// TwinCAT 3 PLC project IAG50cm
// ProjectVersion: 0.10.0
// ProgramVersion: 3.1.4026.12
// libraries:
//   BROTLib, 0.20.0 (BROT)
//   VisuElemBase, * (System)
//   VisuInputs, * (System)
//   Tc2_Math, * (Beckhoff Automation GmbH)
//   Tc2_MC2, * (Beckhoff Automation GmbH)
//   Tc2_MC2_Drive, * (Beckhoff Automation GmbH)
//   Tc2_SerialCom, * (Beckhoff Automation GmbH)
//   Tc2_Standard, * (Beckhoff Automation GmbH)
//   Tc2_System, * (Beckhoff Automation GmbH)
//   Tc2_Utilities, * (Beckhoff Automation GmbH)
//   Tc3_IotBase, * (Beckhoff Automation GmbH)
//   Tc3_IotCommunicator, * (Beckhoff Automation GmbH)
//   Tc3_MC2_AdvancedHoming, * (Beckhoff Automation GmbH)
//   Tc3_Module, * (Beckhoff Automation GmbH)
//   VisuDialogs, * (System)
//   AstroBROT,0.4.3,BROT
//   VisuSymbols,newest,System
// project tree:
//   DUTs/ E_MirrorCoverState.TcDUT, ST_AxisStatus.TcDUT
//   / GlobalTextList.TcGTLO, PlcTask.TcTTO, PlcTask_Fast.TcTTO, Visualization Manager.TcVMO (not stored)
//   GVLs/ GVL_Homing.TcGVL, GVL_Pointing.TcGVL, GVL_Safety.TcGVL, GVL_Serial.TcGVL, Global_Version.TcGVL
//   POUs/CoverControl/ FB_CoverControl.TcPOU
//   POUs/CoverControl/States/ FB_CoverClosingState.TcPOU, FB_CoverIdleState.TcPOU, FB_CoverOpeningState.TcPOU, FB_CoverState.TcPOU, FB_CoverStoppingState.TcPOU, I_CoverState.TcIO
//   POUs/DomeControl/ FB_DomeControl.TcPOU
//   POUs/DomeControl/States/ FB_DomeClosingState.TcPOU, FB_DomeErrorState.TcPOU, FB_DomeHomingState.TcPOU, FB_DomeIdleState.TcPOU, FB_DomeOpeningState.TcPOU, FB_DomeParkingState.TcPOU, FB_DomeStoppingState.TcPOU, FB_DomeState.TcPOU, FB_DomeMovingState.TcPOU, I_DomeState.TcIO
//   POUs/ FB_LatchHome.TcPOU, FB_SafetyHandling.TcPOU, FB_SerialBackground.TcPOU, FB_HomeDropReason.TcPOU, FB_HomeHold.TcPOU, FB_StartRequest.TcPOU, FB_StepDrain.TcPOU, FB_SweepStop.TcPOU, SerialBackground.TcPOU, FB_AxisControl.TcPOU, FB_CabinetControl.TcPOU, FB_FocusControl.TcPOU, FB_HourAngleControl.TcPOU, FB_DeclinationControl.TcPOU, FB_TelescopeControl.TcPOU, MAIN.TcPOU
//   POUs/Functions/ F_HourAngleOffsetOnAxis.TcPOU, F_RoundLREAL.TcPOU, NCError_TO_STRING.TcPOU
//   POUs/PendantControl/ FB_PendantControl.TcPOU
//   POUs/PendantControl/States/ FB_PendantErrorState.TcPOU, FB_PendantPreInitState.TcPOU, FB_PendantSetDECState.TcPOU, FB_PendantSetFocusState.TcPOU, FB_PendantSetHAState.TcPOU, FB_PendantInitState.TcPOU, FB_PendantState.TcPOU, FB_PendantIdleState.TcPOU, I_PendantState.TcIO
//   POUs/Pointing/ FB_PointingModelForward.TcPOU, FB_PointingModelInversion.TcPOU
//   POUs/Testing/ FB_RefMarkerSearch.TcPOU
//   VISUs/ Safety.TcVIS
// real-time tasks:
//   TASK PlcTask: cycle T#10ms, priority 20, ADS port 350
//   TASK VISU_TASK: cycle T#200000us, priority 30, ADS port 351
//   TASK PlcTask_Fast: cycle T#2ms, priority 19, ADS port 352
// motion (NC):
//   TASK NC-Task 1 SAF: cycle T#2ms, priority 4, ADS port 501
//   TASK NC-Task 1 SVB: cycle T#10ms, priority 8, ADS port 511
//   AXIS Declination (id 1)
//     General: UnitName=°
//     Dynamic: Acceleration=3.21148, Deceleration=3.21148, Jerk=4.13844
//     Velo: RefSearch=0.10384, RefSync=0.10384, SlowManual=0.5192, FastManual=3.1152, Fast=10.384, Maximum=10.384
//     TargetPosControl: Range=0.5
//     OtherSettings: AllowMotionCmdToSlave=true
//     encoder EncType=4
//       EncPara: ScaleFactorNumerator=360, ScaleFactorDenominator=36864000, Offset=-23, Inverse=true, MaxCount=#xffffffff
//         Inc: RefMode=2
//     drive DrvType=16
//       DrvPara: MaxCount=#xffffffff, DriveControlDWord=#x00020000
//         Analog: VeloReferenz=11.4224, VeloScale=312, TorqueSetpointScale=10, ScaleFactorActTorque=0.1
//         TimeComp: TaskDelayCycles=1
//     controller CtrType=1
//       CtrPara: PriorControlFactor=1
//         PID: PosKp=3
//         Observer: BandWidth=20
//   AXIS HourAngle (id 2)
//     General: UnitName=°
//     Dynamic: Acceleration=3.6, Deceleration=3.6, Jerk=3.19705
//     Velo: RefSearch=0.10384, RefSync=0.10384, SlowManual=0.5192, FastManual=3.1152, Fast=10.384, Maximum=10.384
//     TargetPosControl: Range=0.5
//     OtherSettings: AllowMotionCmdToSlave=true
//     encoder EncType=4
//       EncPara: ScaleFactorNumerator=360, ScaleFactorDenominator=36864000, Inverse=true, MaxCount=#xffffffff
//         Inc: RefMode=2
//     drive DrvType=16
//       DrvPara: MaxCount=#xffffffff, DriveControlDWord=#x00020000
//         Analog: VeloReferenz=11.4224, VeloScale=312, TorqueSetpointScale=10, ScaleFactorActTorque=0.1
//         TimeComp: TaskDelayCycles=1
//     controller CtrType=1
//       CtrPara: PriorControlFactor=1
//         Observer: BandWidth=20
//   AXIS Focus (id 3)
//     Dynamic: AccelerationMaximum=15, DecelerationMaximum=15, Acceleration=1, Deceleration=1, Jerk=10
//     Velo: RefSearch=0.26997, RefSync=0.26997, SlowManual=0.1, FastManual=1, Fast=26.997, Maximum=2
//     OtherSettings: AllowMotionCmdToSlave=true, PulseDistancePos=1, PulseDistanceNeg=1
//     encoder EncType=19
//       EncPara: ScaleFactorNumerator=3, ScaleFactorDenominator=10485760, Offset=9.78274383544922, MaxCount=#xffffffff, ReferenceSystem=1
//         SoftEndMinControl: Enable=true, Range=1
//         SoftEndMaxControl: Enable=true, Range=17
//     drive DrvType=16
//       DrvPara: MaxCount=#xffffffff, DriveControlDWord=#x00020100
//         Analog: VeloReferenz=29.6967, VeloScale=32, TorqueSetpointScale=10, ScaleFactorActTorque=0.1
//         TimeComp: TaskDelayCycles=1
//     controller CtrType=1
//       CtrPara: PriorControlFactor=1
//         Observer: BandWidth=20
// I/O:
//   DEVICE Device 1 (EtherCAT), AmsNetId 5.146.183.126.2.1
//     Term 1 (EK1200) [EK1200-5000 EtherCAT Power supply (2A E-Bus)]
//       Safety (EL1918) [EL1918, 8Ch. Safety Input 24V, TwinSAFE]
//         modules: Module 2 (FSLOGIC)
//       Safety Out (EL2904) [EL2904, 4 Ch. Safety Output 24V, 0.5A, TwinSAFE]
//         modules: Module 1 (FSOES), Module 2 (DO)
//       Power Status (EL1808) [EL1808 8Ch. Dig. Input 24V, 3ms]
//       HA DEC (ELM7212-9016) [ELM7212-9016 2Ch. Servo Terminal (48 V, 4,5 A RMS, OCT, STO, TwinSAFE Logic)]
//         modules: Module 1 (SAFETY)
//         startup 32785:21 := 0E01 // DRV Motor Settings Ch.1 / Commutation offset
//         startup 32785:27 := 10270000 // DRV Motor Settings Ch.1 / Motor speed limitation
//         startup 32786:19 := 0000 // DRV Brake Settings Ch.1 / Emergency application timeout
//         startup 32784:51 := 0A00 // DRV Amplifier Settings Ch.1 / Stand still window
//         startup 28688:11 := F90C // DRV Outputs Ch.1 / Torque limitation
//         startup 32784:19 := FD00 // DRV Amplifier Settings Ch.1 / Current loop proportional gain
//         startup 32784:18 := 0600 // DRV Amplifier Settings Ch.1 / Current loop integral time
//         startup 32784:21 := 48000000 // DRV Amplifier Settings Ch.1 / Velocity loop proportional gain
//         startup 32784:20 := 96000000 // DRV Amplifier Settings Ch.1 / Velocity loop integral time
//         startup 33041:21 := 0E01 // DRV Motor Settings Ch.2 / Commutation offset
//         startup 33041:27 := 10270000 // DRV Motor Settings Ch.2 / Motor speed limitation
//         startup 33042:19 := 0000 // DRV Brake Settings Ch.2 / Emergency application timeout
//         startup 33040:51 := 0A00 // DRV Amplifier Settings Ch.2 / Stand still window
//         startup 28944:11 := F90C // DRV Outputs Ch.2 / Torque limitation
//         startup 33040:19 := FD00 // DRV Amplifier Settings Ch.2 / Current loop proportional gain
//         startup 33040:18 := 0600 // DRV Amplifier Settings Ch.2 / Current loop integral time
//         startup 33040:21 := 48000000 // DRV Amplifier Settings Ch.2 / Velocity loop proportional gain
//         startup 33040:20 := 96000000 // DRV Amplifier Settings Ch.2 / Velocity loop integral time
//       MirrorCover1 (EL2652) [EL2652 2Ch. Relay Output, CO (230V AC / 30V DC)]
//       MirrorCover2 (EL2652) [EL2652 2Ch. Relay Output, CO (230V AC / 30V DC)]
//       Power (EL9110) [EL9110 Power Supplier with LED (24V, Diagnostics)]
//       Reset 24V (EL2004) [EL2004 4Ch. Dig. Output 24V, 0.5A]
//       FOCUS (ELM7221-9016) [ELM7221-9016 1Ch. Servo Terminal (48 V, 8 A RMS, OCT, STO, TwinSAFE Logic)]
//         modules: Module 1 (SAFETY)
//         startup 32785:21 := 0E01 // DRV Motor Settings Ch.1 / Commutation offset
//         startup 32785:27 := 10270000 // DRV Motor Settings Ch.1 / Motor speed limitation
//         startup 32786:19 := 0000 // DRV Brake Settings Ch.1 / Emergency application timeout
//         startup 32784:51 := 0A00 // DRV Amplifier Settings Ch.1 / Stand still window
//         startup 28688:11 := FC0D // DRV Outputs Ch.1 / Torque limitation
//         startup 32784:19 := FD00 // DRV Amplifier Settings Ch.1 / Current loop proportional gain
//         startup 32784:18 := 0600 // DRV Amplifier Settings Ch.1 / Current loop integral time
//         startup 32784:21 := 47000000 // DRV Amplifier Settings Ch.1 / Velocity loop proportional gain
//         startup 32784:20 := 96000000 // DRV Amplifier Settings Ch.1 / Velocity loop integral time
//       Encoder DEC (EL5021) [EL5021 1Ch. Sin/Cos Encoder]
//       Encoder HA (EL5021) [EL5021 1Ch. Sin/Cos Encoder]
//       Cabinet IN (EL1004) [EL1004 4Ch. Dig. Input 24V, 3ms]
//       Dome Pendant (EL6002) [EL6002 Interface 2Ch. (RS232)]
//       Term 13 (EL9011) [EL9011 End Terminal]
// variable links:
//   Device 1 (EtherCAT) <-> Device 1 (EtherCAT)/Term 1 (EK1200)/FOCUS (ELM7221-9016)
//     Term 1 (EK1200)/Safety (EL1918)/ConnectionOutputs/TwinSafeGroup1.Connection to Term 12 (ELM7221-9016)_3 RxPDO <-> Module 1 (SAFETY)/SAFETY FSoE Connection 1 Send Message/Message_1
//   Device 1 (EtherCAT) <-> Device 1 (EtherCAT)/Term 1 (EK1200)/HA DEC (ELM7212-9016)
//     Term 1 (EK1200)/Safety (EL1918)/ConnectionInputs/TwinSafeGroup1.Connection to Term 4 (ELM7212-9016)_4 TxPDO <-> Module 1 (SAFETY)/SAFETY FSoE Connection 1 Receive Message/Message_1
//     Term 1 (EK1200)/Safety (EL1918)/ConnectionOutputs/TwinSafeGroup1.Connection to Term 4 (ELM7212-9016)_4 RxPDO <-> Module 1 (SAFETY)/SAFETY FSoE Connection 1 Send Message/Message_1
//   Device 1 (EtherCAT) <-> Device 1 (EtherCAT)/Term 1 (EK1200)/Safety (EL1918)
//     Term 1 (EK1200)/FOCUS (ELM7221-9016)/Module 1 (SAFETY)/SAFETY FSoE Connection 1 Receive Message/Message_1 <-> ConnectionInputs/TwinSafeGroup1.Connection to Term 12 (ELM7221-9016)_3 TxPDO
//     Term 1 (EK1200)/Safety Out (EL2904)/Module 1 (FSOES)/RxPDO/FSOE <-> ConnectionInputs/TwinSafeGroup1.EL2904, 4 digital outputs_1_7 TxPDO
//   Device 1 (EtherCAT) <-> Device 1 (EtherCAT)/Term 1 (EK1200)/Safety Out (EL2904)
//     Term 1 (EK1200)/Safety (EL1918)/ConnectionOutputs/TwinSafeGroup1.EL2904, 4 digital outputs_1_7 RxPDO <-> Module 1 (FSOES)/TxPDO/FSOE
//   NC-Task 1 SAF/Axes/Declination <-> Device 1 (EtherCAT)/Term 1 (EK1200)/Encoder DEC (EL5021)
//     Enc/Inputs/In/nDataIn1 <-> ENC Status/Counter value
//     Enc/Inputs/In/nDataIn2 <-> ENC Status/Latch value
//     Enc/Inputs/In/nDcInputTime <-> InfoData/DcInputShift
//     Enc/Inputs/In/nState1 <-> ENC Status/Latch C valid
//     Enc/Inputs/In/nState1 @bit 2 <-> ENC Status/Set counter done
//     Enc/Inputs/In/nState2 @bit 2 <-> ENC Status/Status of input C
//     Enc/Inputs/In/nState2 @bit 5 <-> ENC Status/Sync error
//     Enc/Inputs/In/nState2 @bit 6 <-> ENC Status/TxPDO State
//     Enc/Inputs/In/nState2 @bit 7 <-> ENC Status/TxPDO Toggle
//     Enc/Inputs/In/nState3 @bit 4 <-> ENC Status/Amplitude error
//     Enc/Inputs/In/nState3 @bit 3 <-> ENC Status/Frequency error
//     Enc/Inputs/In/nState4 @bit 1 <-> WcState/InputToggle
//     Enc/Inputs/In/nState4 <-> WcState/WcState
//     Enc/Outputs/Out/nCtrl1 @bit 1 <-> ENC Control/Enable latch C
//     Enc/Outputs/Out/nCtrl1 @bit 2 <-> ENC Control/Set counter
//     Enc/Outputs/Out/nDataOut1 <-> ENC Control/Set counter value
//   NC-Task 1 SAF/Axes/Declination <-> Device 1 (EtherCAT)/Term 1 (EK1200)/HA DEC (ELM7212-9016)
//     Drive/Inputs/In/nDcOutputTime <-> InfoData/DcOutputShift
//     Drive/Inputs/In/nState1 <-> DRV Statusword Channel 1/Statusword
//     Drive/Inputs/In/nState2 <-> DRV Statusword Channel 1/Statusword @bit 8
//     Drive/Inputs/In/nState4 @bit 1 <-> WcState/InputToggle0
//     Drive/Inputs/In/nState4 <-> WcState/WcState0
//     Drive/Outputs/Out/nCtrl1 <-> DRV Controlword Channel 1/Controlword
//     Drive/Outputs/Out/nCtrl2 <-> DRV Controlword Channel 1/Controlword @bit 8
//     Drive/Outputs/Out/nDataOut2 <-> DRV Target velocity Channel 1/Target velocity
//   NC-Task 1 SAF/Axes/Focus <-> Device 1 (EtherCAT)/Term 1 (EK1200)/FOCUS (ELM7221-9016)
//     Drive/Inputs/In/nDataIn1 <-> DRV Following error actual value/Following error actual value
//     Drive/Inputs/In/nDcOutputTime <-> InfoData/DcOutputShift
//     Drive/Inputs/In/nState1 <-> DRV Statusword/Statusword
//     Drive/Inputs/In/nState2 <-> DRV Statusword/Statusword @bit 8
//     Drive/Inputs/In/nState4 @bit 1 <-> WcState/InputToggle0
//     Drive/Inputs/In/nState4 <-> WcState/WcState0
//     Drive/Outputs/Out/nCtrl1 <-> DRV Controlword/Controlword
//     Drive/Outputs/Out/nCtrl2 <-> DRV Controlword/Controlword @bit 8
//     Drive/Outputs/Out/nDataOut1 <-> DRV Target position/Target position
//     Enc/Inputs/In/nDataIn1 <-> FB Position/Position
//     Enc/Inputs/In/nDcInputTime <-> InfoData/DcInputShift
//     Enc/Inputs/In/nState4 @bit 1 <-> WcState/InputToggle0
//     Enc/Inputs/In/nState4 <-> WcState/WcState0
//   NC-Task 1 SAF/Axes/HourAngle <-> Device 1 (EtherCAT)/Term 1 (EK1200)/Encoder HA (EL5021)
//     Enc/Inputs/In/nDataIn1 <-> ENC Status/Counter value
//     Enc/Inputs/In/nDataIn2 <-> ENC Status/Latch value
//     Enc/Inputs/In/nState1 <-> ENC Status/Latch C valid
//     Enc/Inputs/In/nState1 @bit 2 <-> ENC Status/Set counter done
//     Enc/Inputs/In/nState2 @bit 2 <-> ENC Status/Status of input C
//     Enc/Inputs/In/nState2 @bit 5 <-> ENC Status/Sync error
//     Enc/Inputs/In/nState2 @bit 6 <-> ENC Status/TxPDO State
//     Enc/Inputs/In/nState2 @bit 7 <-> ENC Status/TxPDO Toggle
//     Enc/Inputs/In/nState3 @bit 4 <-> ENC Status/Amplitude error
//     Enc/Inputs/In/nState3 @bit 3 <-> ENC Status/Frequency error
//     Enc/Inputs/In/nState4 @bit 1 <-> WcState/InputToggle
//     Enc/Inputs/In/nState4 <-> WcState/WcState
//     Enc/Outputs/Out/nCtrl1 @bit 1 <-> ENC Control/Enable latch C
//     Enc/Outputs/Out/nCtrl1 @bit 2 <-> ENC Control/Set counter
//     Enc/Outputs/Out/nDataOut1 <-> ENC Control/Set counter value
//   NC-Task 1 SAF/Axes/HourAngle <-> Device 1 (EtherCAT)/Term 1 (EK1200)/HA DEC (ELM7212-9016)
//     Drive/Inputs/In/nDcOutputTime <-> InfoData/DcOutputShift
//     Drive/Inputs/In/nState1 <-> DRV Statusword Channel 2/Statusword
//     Drive/Inputs/In/nState2 <-> DRV Statusword Channel 2/Statusword @bit 8
//     Drive/Inputs/In/nState4 @bit 1 <-> WcState/InputToggle0
//     Drive/Inputs/In/nState4 <-> WcState/WcState0
//     Drive/Outputs/Out/nCtrl1 <-> DRV Controlword Channel 2/Controlword
//     Drive/Outputs/Out/nCtrl2 <-> DRV Controlword Channel 2/Controlword @bit 8
//     Drive/Outputs/Out/nDataOut2 <-> DRV Target velocity Channel 2/Target velocity
//   IAG50cm/IAG50cm Instance <-> Device 1 (EtherCAT)/Term 1 (EK1200)/Cabinet IN (EL1004)
//     PlcTask Inputs/MAIN.telescopeControl.fbCabinet.bIMode <-> Channel 1/MAIN.telescopeControl.fbCabinet.bIMode
//     PlcTask Inputs/MAIN.telescopeControl.fbCabinet.bIReset <-> Channel 2/MAIN.telescopeControl.fbCabinet.bIReset
//   IAG50cm/IAG50cm Instance <-> Device 1 (EtherCAT)/Term 1 (EK1200)/Dome Pendant (EL6002)
//     PlcTask_Fast Inputs/SerialBackground.fbDomeSerial.stIn_EL6001/D <-> COM TxPDO-Map Inputs Channel 2/Data In 0
//     PlcTask_Fast Inputs/SerialBackground.fbDomeSerial.stIn_EL6001/D @bit {8..168 step 8} <-> COM TxPDO-Map Inputs Channel 2/Data In {1..21}  (21 links)
//     PlcTask_Fast Inputs/SerialBackground.fbDomeSerial.stIn_EL6001/Status <-> COM TxPDO-Map Inputs Channel 2/Status
//     PlcTask_Fast Inputs/SerialBackground.fbPendantSerial.stIn_EL6001/D <-> COM TxPDO-Map Inputs Channel 1/Data In 0
//     PlcTask_Fast Inputs/SerialBackground.fbPendantSerial.stIn_EL6001/D @bit {8..168 step 8} <-> COM TxPDO-Map Inputs Channel 1/Data In {1..21}  (21 links)
//     PlcTask_Fast Inputs/SerialBackground.fbPendantSerial.stIn_EL6001/Status <-> COM TxPDO-Map Inputs Channel 1/Status
//     PlcTask_Fast Outputs/SerialBackground.fbDomeSerial.stOut_EL6001/Ctrl <-> COM RxPDO-Map Outputs Channel 2/Ctrl
//     PlcTask_Fast Outputs/SerialBackground.fbDomeSerial.stOut_EL6001/D <-> COM RxPDO-Map Outputs Channel 2/Data Out 0
//     PlcTask_Fast Outputs/SerialBackground.fbDomeSerial.stOut_EL6001/D @bit {8..168 step 8} <-> COM RxPDO-Map Outputs Channel 2/Data Out {1..21}  (21 links)
//     PlcTask_Fast Outputs/SerialBackground.fbPendantSerial.stOut_EL6001/Ctrl <-> COM RxPDO-Map Outputs Channel 1/Ctrl
//     PlcTask_Fast Outputs/SerialBackground.fbPendantSerial.stOut_EL6001/D <-> COM RxPDO-Map Outputs Channel 1/Data Out 0
//     PlcTask_Fast Outputs/SerialBackground.fbPendantSerial.stOut_EL6001/D @bit {8..168 step 8} <-> COM RxPDO-Map Outputs Channel 1/Data Out {1..21}  (21 links)
//   IAG50cm/IAG50cm Instance <-> Device 1 (EtherCAT)/Term 1 (EK1200)/FOCUS (ELM7221-9016)
//     PlcTask Outputs/GVL_Safety.ErrAck <-> Module 1 (SAFETY)/SAFETY Standard Outputdata/Standard In Var 3
//     PlcTask Outputs/GVL_Safety.Run <-> Module 1 (SAFETY)/SAFETY Standard Outputdata/Standard In Var 2
//   IAG50cm/IAG50cm Instance <-> Device 1 (EtherCAT)/Term 1 (EK1200)/HA DEC (ELM7212-9016)
//     PlcTask Outputs/GVL_Safety.ErrAck <-> Module 1 (SAFETY)/SAFETY Standard Outputdata/Standard In Var 3
//     PlcTask Outputs/GVL_Safety.Run <-> Module 1 (SAFETY)/SAFETY Standard Outputdata/Standard In Var 2
//   IAG50cm/IAG50cm Instance <-> Device 1 (EtherCAT)/Term 1 (EK1200)/MirrorCover1 (EL2652)
//     PlcTask Outputs/MAIN.coverControl.bMotor1RelaisA <-> Channel 1/Output
//     PlcTask Outputs/MAIN.coverControl.bMotor1RelaisB <-> Channel 2/Output
//   IAG50cm/IAG50cm Instance <-> Device 1 (EtherCAT)/Term 1 (EK1200)/MirrorCover2 (EL2652)
//     PlcTask Outputs/MAIN.coverControl.bMotor2RelaisA <-> Channel 1/Output
//     PlcTask Outputs/MAIN.coverControl.bMotor2RelaisB <-> Channel 2/Output
//   IAG50cm/IAG50cm Instance <-> Device 1 (EtherCAT)/Term 1 (EK1200)/Power Status (EL1808)
//     PlcTask Inputs/MAIN.telescopeControl.fbCabinet.bAuxiliaryContact24V <-> Channel 1/Input
//     PlcTask Inputs/MAIN.telescopeControl.fbCabinet.bAuxiliaryContact48V <-> Channel 2/Input
//     PlcTask Inputs/MAIN.telescopeControl.fbCabinet.bAuxiliaryContactFOCUS <-> Channel 4/Input
//     PlcTask Inputs/MAIN.telescopeControl.fbCabinet.bAuxiliaryContactHADEC <-> Channel 3/Input
//     PlcTask Inputs/MAIN.telescopeControl.fbCabinet.bCollectiveReport24VFuse <-> Channel 6/Input
//     PlcTask Inputs/MAIN.telescopeControl.fbCabinet.bState24VFuse <-> Channel 5/Input
//   IAG50cm/IAG50cm Instance <-> Device 1 (EtherCAT)/Term 1 (EK1200)/Reset 24V (EL2004)
//     PlcTask Outputs/MAIN.telescopeControl.fbCabinet.bOErrorLED <-> Channel 2/MAIN.telescopeControl.fbCabinet.bOErrorLED
//   IAG50cm/IAG50cm Instance <-> Device 1 (EtherCAT)/Term 1 (EK1200)/Safety (EL1918)
//     PlcTask Inputs/MAIN.safetyHandling.stInfoEStop1 <-> Function Block Info Data/TwinSafeGroup1.SS1.FBMon1 Info Data
//     PlcTask Inputs/MAIN.safetyHandling.stInfoGroup1 <-> TwinSAFE Group Info Data/TwinSafeGroup1 Info Data
//     PlcTask Outputs/GVL_Safety.ErrAck <-> StandardOutputs/TwinSafeGroup1.ErrorAcknowledgement_2
//     PlcTask Outputs/GVL_Safety.Restart <-> StandardOutputs/TwinSafeGroup1.Restart_6
//     PlcTask Outputs/GVL_Safety.Run <-> StandardOutputs/TwinSafeGroup1.Run_1
//   IAG50cm/IAG50cm Instance <-> NC-Task 1 SAF/Axes/Declination
//     PlcTask Inputs/MAIN.decControl.axisRef.NcToPlc <-> Outputs/ToPlc
//     PlcTask Outputs/MAIN.decControl.axisRef.PlcToNc <-> Inputs/FromPlc
//   IAG50cm/IAG50cm Instance <-> NC-Task 1 SAF/Axes/Focus
//     PlcTask Inputs/MAIN.focusControl.axisRef.NcToPlc <-> Outputs/ToPlc
//     PlcTask Outputs/MAIN.focusControl.axisRef.PlcToNc <-> Inputs/FromPlc
//   IAG50cm/IAG50cm Instance <-> NC-Task 1 SAF/Axes/HourAngle
//     PlcTask Inputs/MAIN.haControl.axisRef.NcToPlc <-> Outputs/ToPlc
//     PlcTask Outputs/MAIN.haControl.axisRef.PlcToNc <-> Inputs/FromPlc

CONFIGURATION IAG50cm
    RESOURCE PLC ON TwinCAT3
        TASK PlcTask(INTERVAL := T#10ms, PRIORITY := 20);
        TASK PlcTask_Fast(INTERVAL := T#2ms, PRIORITY := 19);
        PROGRAM MAIN WITH PlcTask : MAIN;
        PROGRAM SerialBackground WITH PlcTask_Fast : SerialBackground;
    END_RESOURCE
END_CONFIGURATION

// ---- DUTs/E_MirrorCoverState.TcDUT
{attribute 'qualified_only'}
{attribute 'strict'}
//{attribute 'to_string'}
TYPE E_MirrorCoverState :
(
	closing := 0,
	opening := 1,
	stopped := 2,
	closed	:= 3,
	open	:= 4,
	error := 5,
	unknown := 6
);
END_TYPE

// ---- DUTs/ST_AxisStatus.TcDUT
// Plan step 3.2: the feedback of one axis (FB_Axis outputs) as read once per scan by FB_TelescopeControl._ReadAxes. Same struct as
// MONETcommon's (it moves to BROTLib in step 4). The axes' outputs do not change while the telescope body runs, so reading them into
// one struct is the same as reading fbAxis.* at every use.
TYPE ST_AxisStatus :
STRUCT
	bStandStill		: BOOL;
	bStopDone		: BOOL;
	bInMotion		: BOOL;
	bInRamp			: BOOL;
	bHoming			: BOOL;
	bStopping		: BOOL;
	bBusy			: BOOL;
	bTracking		: BOOL;
END_STRUCT
END_TYPE

// ---- GVLs/GVL_Homing.TcGVL
{attribute 'qualified_only'}
VAR_GLOBAL
	// #113: how FB_LatchHome ends the calibration sweep after a stop. Test switch, written over ADS (GVL_Homing.nAbortMode),
	// so the approaches can be tried one after the other without a new activation. Not persistent.
	//   0: as before (MC_AbortHoming into the running step: never completes, 4F000001 after 10 s)
	//   1: no MC_AbortHoming while a step block is Busy, the axis is reset instead (reset=1 clears HomingBusy)
	//   2: the Busy reference step keeps its Execute while MC_AbortHoming runs
	//   3: MC_AbortHoming with DisableDriveAccess FALSE
	nAbortMode		: INT := 1;
END_VAR

// ---- GVLs/GVL_Pointing.TcGVL
VAR_GLOBAL
	(* values of the pointing model
	Hour Angle	: tau
	Declination	: dec
	*)

	(*
	 pointing from: 21.01.2026 136 points (from Lukas Melzig)
	RMS Ha:  17.69244750276253
	RMS Dec:  13.468555776826959
	*)
	C_mAl_tau	: LREAL := 0.01687078;
	C_mEl_tau	: LREAL := -0.02608578;
	C_Coll_tau	: LREAL := 0.29826615;
	C_Refr_tau	: LREAL := -0.00759962;
	C_Enc_tau	: LREAL := 0.00108764;
	C_Flex_tau	: LREAL := -0.02462705;
	C_NP_tau	: LREAL := 0.02128217;
	
	C_mAl_dec	: LREAL := 0.01606325;
	C_mEl_dec	: LREAL := -0.05749048;
	C_Coll_dec	: LREAL := -0.17376101;
	C_Refr_dec	: LREAL := 0.01678090;
	C_Flex_dec	: LREAL := -0.01915146;
END_VAR

// ---- GVLs/GVL_Safety.TcGVL
{attribute 'qualified_only'}
VAR_GLOBAL
	// Run/Stop Safety
	Run			AT%Q*:	BOOL;
	// Restart Safety
	Restart		AT%Q*:	BOOL;
	// Error Acknowledgement 
	ErrAck		AT%Q*:	BOOL;

END_VAR

// ---- GVLs/GVL_Serial.TcGVL
VAR_GLOBAL
	RxBufferDome			: ComBuffer;	(* Receive data buffer; used with all receive function blocks *)
	TxBufferDome			: ComBuffer;	(* Transmit data buffer; used with all receive function blocks *)
	
	RxBufferPendant			: ComBuffer;	(* Receive data buffer; used with all receive function blocks *)
	TxBufferPendant			: ComBuffer;	(* Transmit data buffer; used with all receive function blocks *)
END_VAR

// ---- GVLs/Global_Version.TcGVL
{attribute 'qualified_only'}
VAR_GLOBAL CONSTANT
	// Mirrors Beckhoff's own Global_Version.stLibVersion_* pattern (see ST_LibVersion),
	// which only covers Tc2_*/Tc3_* library references, not custom ones -- until now: this
	// GVL uses Beckhoff's own naming exactly, so it merges into a consumer's Global_Version.
	// Kept in sync with <ProjectVersion> in IAG50cm.plcproj at release time.
	stLibVersion_IAG50cm : ST_LibVersion := (
		iMajor := 0,
		iMinor := 10,
		iBuild := 0,
		iRevision := 0,
		nFlags := 1,
		sVersion := '0.10.0'
	);
END_VAR

// ---- POUs/CoverControl/States/I_CoverState.TcIO
INTERFACE I_CoverState

METHOD CloseCommand : BOOL
VAR_INPUT
END_VAR
END_METHOD

METHOD OpenCommand : BOOL
VAR_INPUT
END_VAR
END_METHOD

METHOD RunState : BOOL
VAR_INPUT
END_VAR
END_METHOD

METHOD StopCommand : BOOL
VAR_INPUT
END_VAR
END_METHOD

METHOD SuccessfulFinished : BOOL
VAR_INPUT
END_VAR
END_METHOD

END_INTERFACE

// ---- POUs/DomeControl/States/I_DomeState.TcIO
INTERFACE I_DomeState


METHOD CloseCommand : BOOL
END_METHOD


METHOD FoundError : BOOL
END_METHOD


METHOD HomeCommand : BOOL
END_METHOD


METHOD MoveCommand : BOOL
END_METHOD


METHOD OpenCommand : BOOL
END_METHOD


METHOD ParkCommand : BOOL
END_METHOD


METHOD ResetCommand : BOOL
END_METHOD

METHOD RunState : BOOL
VAR_INPUT
END_VAR
END_METHOD


PROPERTY StateID : STRING
GET
END_GET
END_PROPERTY


METHOD StopCommand : BOOL
END_METHOD


METHOD SuccessfulFinished : BOOL
END_METHOD

END_INTERFACE

// ---- POUs/PendantControl/States/I_PendantState.TcIO
INTERFACE I_PendantState

METHOD DecCommand : BOOL
VAR_INPUT
END_VAR
END_METHOD

METHOD FocusCommand : BOOL
VAR_INPUT
END_VAR
END_METHOD

METHOD FoundError : BOOL
VAR_INPUT
END_VAR
END_METHOD

METHOD HaCommand : BOOL
VAR_INPUT
END_VAR
END_METHOD

METHOD InitCommand : BOOL
VAR_INPUT
END_VAR
END_METHOD

METHOD ResetCommand : BOOL
VAR_INPUT
END_VAR
END_METHOD

METHOD RunState : BOOL
VAR_INPUT
END_VAR
END_METHOD

PROPERTY StateID : STRING
GET
END_GET
END_PROPERTY

METHOD Timeout : BOOL
VAR_INPUT
END_VAR
END_METHOD

METHOD ToIdle : BOOL
VAR_INPUT
END_VAR
END_METHOD

END_INTERFACE

// ---- POUs/MAIN.TcPOU
PROGRAM MAIN
VAR
	comm			: FB_Comm_MQTT_Influx;
	coverControl	: FB_CoverControl(comm := comm);
	focusControl	: FB_FocusControl(comm:=comm);
	haControl		: FB_HourAngleControl(comm:=comm);
	decControl		: FB_DeclinationControl(comm:=comm);
	telescopeControl: FB_TelescopeControl(comm := comm);
	domeControl		: FB_DomeControl(comm := comm);
	pendantControl 	: FB_PendantControl(comm:=comm);
	safetyHandling	: FB_SafetyHandling(comm:=comm);
	rtrigStartUpDone: R_TRIG;
	//search			: FB_RefMarkerSearch(); // use for searching for the Heideinhain encoder reference markers

	
END_VAR
VAR CONSTANT
	telescopeConfig		: ST_TelescopeConfig := (longitude := 9.9452433, latitude := 51.5592378, altitude := 100.0, 
													houranglePark := 0.0, declinationPark := 52.0, focusPark:= 16.3,
													hourangleHome := 0.0, declinationHome := 52.0, focusHome:= 16.3,
													name := 'Emmy Noether', diameter := 0.5, cabinet := 'Beckhoff', manufacturer := '???',
													mountOptions := 'HA-DEC', mount := 'HA_DEC');
END_VAR

//search(Enable:=TRUE); // use for reference marker search

domeControl(ipTelescope	:= telescopeControl);

pendantControl(
	ipTelescope	:= telescopeControl,
	ipFocus		:= focusControl);

coverControl(
	Delta := T#5S,
	TimeToCycle := T#15S,
	bEmergency := safetyHandling.estop);	// previous cycle's value, see bEstopTriggered below (#15)
	
focusControl(
	fVelocity:=1);
	
haControl();
decControl();
telescopeControl(
	fbHourAngle		:= haControl,
	fbDeclination	:= decControl,
	fbFocus			:= focusControl,
	fbDome			:= domeControl,
	fbCovers		:= coverControl,
	telescopeConfig	:= telescopeConfig,
	// was never wired, so STATUS.GLOBAL never reported the E-stop (BROTLib#10). safetyHandling runs below, so
	// this is the previous cycle's value; the drives are cut by the safety circuit regardless.
	bEstopTriggered	:= safetyHandling.estop,
	bSafetyAckPending	:= safetyHandling.ackPending,	// previous cycle, like bEstopTriggered (#59)
);

//Safety
// #11: a telescope reset (cabinet key or the reset command, only fires with an error or a pending acknowledge after an E-stop, #59) also gives the safety
// acknowledge, so the drives leave STO without the VISU
IF telescopeControl.bSafetyAckRequest THEN
	telescopeControl.bSafetyAckRequest := FALSE;
	safetyHandling.Acknowledge();
END_IF
safetyHandling();
// #103: one axis reset pass once the safety start-up is done (the start-up only acknowledges the drives)
rtrigStartUpDone(CLK := safetyHandling.bStartUpDone);
IF rtrigStartUpDone.Q THEN
	telescopeControl.bStartupAxisReset := TRUE;
END_IF

// Comm
comm(	
	sHostName			:= '169.254.149.100',
    nHostPort  			:= 1883,
    nKeepAlive  		:= 10,
	sTopicSub  		 	:= '50cm/Telescope/SET',
	sTopicPublish		:= '50cm/Telemetry',
	sTopicLog			:= '50cm/Log',
	Telescope			:= telescopeControl,
	RaDecTelescope		:= telescopeControl,
	Focus				:= focusControl,
	Dome				:= domeControl,
	MirrorCovers		:= coverControl,
);

END_PROGRAM

// ---- POUs/CoverControl/FB_CoverControl.TcPOU
FUNCTION_BLOCK FB_CoverControl IMPLEMENTS I_MirrorCovers
VAR_INPUT
	Delta		: TIME := T#5S;		// Time difference between both covers opening (and closing)
	TimeToCycle	: TIME := T#15S;	// Time for one motor to fully open/close
	// TRUE while the E-stop is triggered (MAIN: safetyHandling.estop): moving covers stop, open/close requests
	// are dropped (#15)
	bEmergency	: BOOL;
END_VAR
VAR_OUTPUT
END_VAR
VAR
	bOpen		: BOOL;
	bClose		: BOOL;
	bStop		: BOOL;
	// State
	fbCoverIdleState : FB_CoverIdleState(THIS);
	fbCoverOpeningState : FB_CoverOpeningState(THIS);
	fbCoverStoppingState : FB_CoverStoppingState(THIS);
	fbCoverClosingState : FB_CoverClosingState(THIS);
	
	ipState		: I_CoverState := fbCoverIdleState;
	// #111: the PLC cannot know the position of the covers after a start (activation, Reset Cold), so it starts with
	// "unknown" instead of assuming "closed". The first open or close cycle that completes sets the real end position.
	eCoverState	: E_MirrorCoverState := E_MirrorCoverState.unknown;
	// #71: TRUE only once an open or close cycle has completed since the PLC start. Until then the position is
	// unknown (the covers may be open after a restart), so a request is only ignored once the position is confirmed.
	bEndPositionConfirmed : BOOL := FALSE;
	bRequestIgnored : BOOL;
	// Trigger
	rtrigOpen		: R_TRIG;
	rtrigClose		: R_TRIG;
	rtrigStop		: R_TRIG;
	// Comm
	fbComm			: I_Comm;
	tonComm 		: TON := (PT:=T#5S);
	fbCoverOpenEvent:	FB_EventLog;
	fbCoverClosedEvent: FB_EventLog;
	fbCoverEmergencyEvent: FB_EventLog;
	fbCoverIgnoredEvent: FB_EventLog;
	// Motor relais
	bMotor1RelaisA	AT%Q*	: BOOL := FALSE;
	bMotor1RelaisB	AT%Q*	: BOOL := FALSE;
	
	bMotor2RelaisA	AT%Q*	: BOOL := FALSE;
	bMotor2RelaisB	AT%Q*	: BOOL := FALSE;
END_VAR

rtrigOpen(CLK := bOpen);
rtrigClose(CLK := bClose);
rtrigStop(CLK := bStop);
bRequestIgnored := FALSE;

IF bEmergency THEN
	// requests made during the E-stop are dropped (flags cleared below, #15)
	// stop only moving covers, so that closed/open covers keep their known state
	IF eCoverState = E_MirrorCoverState.opening OR eCoverState = E_MirrorCoverState.closing THEN
		ipState.StopCommand();
	END_IF
ELSE
	IF rtrigStop.Q THEN
		ipState.StopCommand();
	END_IF

	// #71: a request for the position the covers are confirmed to be in does nothing (it ran a full 20 s cycle)
	IF rtrigClose.Q THEN
		IF eCoverState = E_MirrorCoverState.closed AND bEndPositionConfirmed THEN
			bRequestIgnored := TRUE;
		ELSE
			ipState.CloseCommand();
		END_IF
	END_IF

	IF rtrigOpen.Q THEN
		IF eCoverState = E_MirrorCoverState.open AND bEndPositionConfirmed THEN
			bRequestIgnored := TRUE;
		ELSE
			ipState.OpenCommand();
		END_IF
	END_IF
END_IF

// #66: requests are one-shot. They are consumed in this scan whether they produced an edge or not, so a caller that
// repeats a request every scan (the park, stage 80) cannot leave a flag TRUE: left set, it would block the rising
// edge of every later request.
bOpen := FALSE;
bClose := FALSE;
bStop := FALSE;

ipState.RunState();

// send telemetry
tonComm(IN:=TRUE);
IF tonComm.Q THEN // publish new payload every second
	tonComm(IN:=FALSE);
	THIS^._SendTelemetry();	
END_IF


fbCoverOpenEvent(
	Trigger := eCoverState = E_MirrorCoverState.open,
	Level := ADSLOG_MSGTYPE_HINT,
	OnMessage := 'Mirror cover is open.',
	comm:= fbComm);
fbCoverClosedEvent(
	Trigger := eCoverState = E_MirrorCoverState.closed,
	Level := ADSLOG_MSGTYPE_HINT,
	OnMessage := 'Mirror cover is closed.',
	comm:= fbComm);
fbCoverIgnoredEvent(
	Trigger := bRequestIgnored,
	Level := ADSLOG_MSGTYPE_HINT,
	OnMessage := 'Mirror cover already in the requested end position, request ignored.',
	comm:= fbComm);
fbCoverEmergencyEvent(
	Trigger := bEmergency,
	Level := ADSLOG_MSGTYPE_WARN,
	OnMessage := 'Mirror cover: E-stop, covers stopped and commands ignored.',
	comm:= fbComm);

PROPERTY _CoverState : E_MirrorCoverState
SET
eCoverState := _CoverState;
bEndPositionConfirmed := (_CoverState = E_MirrorCoverState.closed OR _CoverState = E_MirrorCoverState.open);
END_SET
END_PROPERTY

PROPERTY _Motor1RelaisA : BOOL
SET
bMotor1RelaisA := _Motor1RelaisA;
END_SET
END_PROPERTY

PROPERTY _Motor1RelaisB : BOOL
SET
bMotor1RelaisB := _Motor1RelaisB;
END_SET
END_PROPERTY

PROPERTY _Motor2RelaisA : BOOL
SET
bMotor2RelaisA := _Motor2RelaisA;
END_SET
END_PROPERTY

PROPERTY _Motor2RelaisB : BOOL
SET
bMotor2RelaisB := _Motor2RelaisB;
END_SET
END_PROPERTY

METHOD _SendTelemetry : BOOL
VAR_INPUT
END_VAR
IF eCoverState = E_MirrorCoverState.closed THEN
	fbComm.PublishLREAL('telescope', 'dome', 'AUXILIARY.COVER.REALPOS', 0.0);
ELSIF eCoverState = E_MirrorCoverState.open THEN
	fbComm.PublishLREAL('telescope', 'dome', 'AUXILIARY.COVER.REALPOS', 1.0);
ELSE
	// moving, stopped or unknown (#111): not at an end position
	fbComm.PublishLREAL('telescope', 'dome', 'AUXILIARY.COVER.REALPOS', 0.5);
END_IF
END_METHOD

METHOD Close : BOOL
VAR_INPUT
END_VAR
bClose := TRUE;
END_METHOD

PROPERTY Closed : BOOL
GET
IF THIS^.CoverState = E_MirrorCoverState.closed THEN
	Closed := TRUE;
ELSE
	Closed := FALSE;
END_IF
END_GET
END_PROPERTY

PROPERTY CoverState : E_MirrorCoverState
GET
CoverState := eCoverState;
END_GET
END_PROPERTY

PROPERTY Error : BOOL
GET
Error := FALSE;
END_GET
END_PROPERTY

//FB_Init is always available implicitly and it is used primarily for initialization.
//The return value is not evaluated. For a specific influence, you can also declare the
//methods explicitly and provide additional code there with the standard initialization
//code. You can evaluate the return value.
METHOD FB_Init: BOOL
VAR_INPUT
    bInitRetains	: BOOL; // TRUE: the retain variables are initialized (reset warm / reset cold)
    bInCopyCode		: BOOL;  // TRUE: the instance will be copied to the copy code afterward (online change)
	comm			: I_Comm;
END_VAR
THIS^.fbComm 				:= comm;
END_METHOD

METHOD Open : BOOL
VAR_INPUT
END_VAR
bOpen := TRUE;
END_METHOD

PROPERTY Opened : BOOL
GET
IF THIS^.CoverState = E_MirrorCoverState.open THEN
	Opened := TRUE;
ELSE
	Opened := FALSE;
END_IF
END_GET
END_PROPERTY

METHOD Reset : BOOL
VAR_INPUT
END_VAR
END_METHOD

METHOD SetState : BOOL
VAR_INPUT
	newState :I_CoverState;
END_VAR
THIS^.ipState := newState;
END_METHOD

METHOD Stop : BOOL
VAR_INPUT
END_VAR
bStop := TRUE;
END_METHOD

END_FUNCTION_BLOCK

// ---- POUs/CoverControl/States/FB_CoverIdleState.TcPOU
FUNCTION_BLOCK FB_CoverIdleState EXTENDS FB_CoverState
VAR_INPUT
END_VAR
VAR_OUTPUT
END_VAR
VAR
END_VAR

METHOD CloseCommand : BOOL
pCover^.SetState(pCover^.fbCoverClosingState);
END_METHOD

METHOD OpenCommand : BOOL
pCover^.SetState(pCover^.fbCoverOpeningState);
END_METHOD

METHOD StopCommand : BOOL
pCover^.SetState(pCover^.fbCoverStoppingState);
END_METHOD

END_FUNCTION_BLOCK

// ---- POUs/CoverControl/States/FB_CoverState.TcPOU
FUNCTION_BLOCK FB_CoverState IMPLEMENTS I_CoverState
VAR_INPUT
END_VAR
VAR_OUTPUT
END_VAR
VAR
	pCover : POINTER TO FB_CoverControl;
END_VAR

{warning 'add method implementation '}
METHOD CloseCommand : BOOL
END_METHOD

METHOD FB_init : BOOL
VAR_INPUT
	bInitRetains : BOOL; // if TRUE, the retain variables are initialized (warm start / cold start)
	bInCopyCode : BOOL;  // if TRUE, the instance afterwards gets moved into the copy code (online change)
	pCover : POINTER TO FB_CoverControl;
END_VAR
THIS^.pCover := pCover;
END_METHOD

{warning 'add method implementation '}
METHOD OpenCommand : BOOL
END_METHOD

{warning 'add method implementation '}
METHOD RunState : BOOL
END_METHOD

{warning 'add method implementation '}
METHOD StopCommand : BOOL
END_METHOD

{warning 'add method implementation '}
METHOD SuccessfulFinished : BOOL
END_METHOD

END_FUNCTION_BLOCK

// ---- POUs/CoverControl/States/FB_CoverOpeningState.TcPOU
FUNCTION_BLOCK FB_CoverOpeningState EXTENDS FB_CoverState
VAR
	nStage			: UINT:= 0;
	tonDelta		: TON;		// PT is taken from pCover^.Delta at the start of each cycle (#76)
	tonFullCycle	: TON;		// PT is taken from pCover^.TimeToCycle at the start of each cycle (#76)
END_VAR

METHOD CloseCommand : BOOL
nStage := 0;
tonDelta(IN:=FALSE);
tonFullCycle(IN:=FALSE);
pCover^.SetState(pCover^.fbCoverClosingState);
END_METHOD

METHOD RunState : BOOL
tonDelta();
tonFullCycle();
CASE nStage OF
	0:
		// #76: the cycle times were only read once, by the declaration initialisers, so the inputs of FB_CoverControl
		// never reached the timers. Take them at the start of each cycle (not every scan: a change mid-cycle must not
		// end it early).
		tonDelta.PT := pCover^.Delta;
		IF pCover^.TimeToCycle > T#0S THEN
			tonFullCycle.PT := pCover^.TimeToCycle;
		ELSE
			tonFullCycle.PT := T#15S;	// 0 would declare the end position after one scan
		END_IF
		pCover^._CoverState := E_MirrorCoverState.opening;
		tonDelta.IN:=TRUE;
		nStage := 1;
	1:
		// Open Motor 1
		pCover^._Motor1RelaisA := TRUE;
		pCover^._Motor1RelaisB := FALSE;
		// Stop Motor 2
		pCover^._Motor2RelaisA := FALSE;
		pCover^._Motor2RelaisB := FALSE;
		nStage := 2;
	2:
		IF tonDelta.Q THEN
			tonDelta.IN:=FALSE;
			nStage:=3;
		END_IF 
	3:
		// Open Motor 2
		pCover^._Motor2RelaisA := TRUE;
		pCover^._Motor2RelaisB := FALSE;
		tonFullCycle.IN:=TRUE;
		nStage := 4;
	4:
		IF tonFullCycle.Q THEN
			tonFullCycle.IN:=FALSE;
			THIS^.SuccessfulFinished();
		END_IF 
END_CASE
END_METHOD

METHOD StopCommand : BOOL
nStage := 0;
tonDelta(IN:=FALSE);
tonFullCycle(IN:=FALSE);
pCover^.SetState(pCover^.fbCoverStoppingState);
END_METHOD

METHOD SuccessfulFinished : BOOL
nStage := 0;
tonDelta(IN:=FALSE);
tonFullCycle(IN:=FALSE);
// #71: release the relays at the end position (limit switches cut the motors, the covers are self-locking)
pCover^._Motor1RelaisA := FALSE;
pCover^._Motor1RelaisB := FALSE;
pCover^._Motor2RelaisA := FALSE;
pCover^._Motor2RelaisB := FALSE;
pCover^._CoverState := E_MirrorCoverState.open;
pCover^.SetState(pCover^.fbCoverIdleState);
END_METHOD

END_FUNCTION_BLOCK

// ---- POUs/CoverControl/States/FB_CoverStoppingState.TcPOU
FUNCTION_BLOCK FB_CoverStoppingState EXTENDS FB_CoverState
VAR_INPUT
END_VAR
VAR_OUTPUT
END_VAR
VAR
END_VAR

METHOD RunState : BOOL
// Stop Motor 1
pCover^._Motor1RelaisA := FALSE;
pCover^._Motor1RelaisB := FALSE;
// Stop Motor 2
pCover^._Motor2RelaisA := FALSE;
pCover^._Motor2RelaisB := FALSE;
THIS^.SuccessfulFinished();
END_METHOD

METHOD SuccessfulFinished : BOOL
pCover^._CoverState := E_MirrorCoverState.stopped;
pCover^.SetState(pCover^.fbCoverIdleState);
END_METHOD

END_FUNCTION_BLOCK

// ---- POUs/CoverControl/States/FB_CoverClosingState.TcPOU
FUNCTION_BLOCK FB_CoverClosingState EXTENDS FB_CoverState
VAR
	nStage			: UINT:= 0;
	tonDelta		: TON;		// PT is taken from pCover^.Delta at the start of each cycle (#76)
	tonFullCycle	: TON;		// PT is taken from pCover^.TimeToCycle at the start of each cycle (#76)
END_VAR

METHOD OpenCommand : BOOL
nStage := 0;
tonDelta(IN:=FALSE);
tonFullCycle(IN:=FALSE);
pCover^.SetState(pCover^.fbCoverOpeningState);
END_METHOD

METHOD RunState : BOOL
tonDelta();
tonFullCycle();
CASE nStage OF
	0:
		// #76: the cycle times were only read once, by the declaration initialisers, so the inputs of FB_CoverControl
		// never reached the timers. Take them at the start of each cycle (not every scan: a change mid-cycle must not
		// end it early).
		tonDelta.PT := pCover^.Delta;
		IF pCover^.TimeToCycle > T#0S THEN
			tonFullCycle.PT := pCover^.TimeToCycle;
		ELSE
			tonFullCycle.PT := T#15S;	// 0 would declare the end position after one scan
		END_IF
		pCover^._CoverState := E_MirrorCoverState.closing;
		tonDelta.IN := TRUE;
		nStage := 1;
	1:
		// Stop Motor 1
		pCover^._Motor1RelaisA := FALSE;
		pCover^._Motor1RelaisB := FALSE;
		// Close Motor 2
		pCover^._Motor2RelaisA := FALSE;
		pCover^._Motor2RelaisB := TRUE;
		nStage := 2;
	2:
		IF tonDelta.Q THEN
			tonDelta.IN := FALSE;
			nStage:=3;
		END_IF 
	3:
		// Close Motor 1
		pCover^._Motor1RelaisA := FALSE;
		pCover^._Motor1RelaisB := TRUE;
		tonFullCycle.IN:=TRUE;
		nStage := 4;
	4:
		IF tonFullCycle.Q THEN
			tonFullCycle.IN := FALSE;
			THIS^.SuccessfulFinished();
		END_IF 
END_CASE
END_METHOD

METHOD StopCommand : BOOL
nStage := 0;
tonDelta(IN:=FALSE);
tonFullCycle(IN:=FALSE);
pCover^.SetState(pCover^.fbCoverStoppingState);
END_METHOD

METHOD SuccessfulFinished : BOOL
nStage := 0;
tonDelta(IN:=FALSE);
tonFullCycle(IN:=FALSE);
// #71: release the relays at the end position (limit switches cut the motors, the covers are self-locking)
pCover^._Motor1RelaisA := FALSE;
pCover^._Motor1RelaisB := FALSE;
pCover^._Motor2RelaisA := FALSE;
pCover^._Motor2RelaisB := FALSE;
pCover^._CoverState := E_MirrorCoverState.closed;
pCover^.SetState(pCover^.fbCoverIdleState);
END_METHOD

END_FUNCTION_BLOCK

// ---- POUs/FB_FocusControl.TcPOU
FUNCTION_BLOCK FB_FocusControl EXTENDS FB_AxisControl IMPLEMENTS I_Focus
VAR_INPUT
	fMinPosition		: LREAL := 1.0;			// minimum Position
	fMaxPosition		: LREAL := 17.0;		// maximum Position
	fTolerance			: LREAL := 0.005;
END_VAR
VAR
	mqttTimer 			: TON := (PT:=T#5S);
	fbFollower			: BROTLib.FB_MoveFollower;	// starts, re-targets and holds the move to fPosition (MONETcommon#122)
	bHoldOnStop			: BOOL;		// Stop() was called: the target becomes the position reached at StopDone
END_VAR

// limit to sane positions
fPosition := LIMIT(fMinPosition, fPosition, fMaxPosition);


IF bEnable AND NOT fbAxis.Calibrated THEN
	THIS^.HomeAxis := TRUE;		// starts _StartHoming on FALSE -> TRUE
END_IF

// a new target during a move restarts it, MoveDone, abort, error and stop end it (MONETcommon#122); the inputs are
// what fbAxis reported in its last call. The enable comes from the telescope, so bNeedEnable is not used.
fbFollower(
	fTarget		:= fPosition,
	fActual		:= fActualPosition,
	fTolerance	:= fTolerance,
	bActive		:= fbAxis.Calibrated,
	bReady		:= fbAxis.Ready AND NOT fbAxis.MoveDone,
	bMoveDone	:= fbAxis.MoveDone,
	bAborted	:= fbAxis.CommandAborted,
	bError		:= bError,
	bStopDone	:= fbAxis.StopDone);

// Stop(): hold the position reached when the stop is done
IF bHoldOnStop AND (fbAxis.StopDone OR fbAxis.StandStill) THEN
	bHoldOnStop := FALSE;
	IF fbAxis.Calibrated THEN
		fPosition := fActualPosition;
	END_IF
END_IF

// after an error a reset must not resume the old move by itself
IF bError AND fbAxis.Calibrated THEN
	fPosition := fActualPosition;
END_IF

IF fbAxis.Calibrated THEN
	bHomeAxis := FALSE;
	bCalibrated := fbAxis.Calibrated;
	// MoveTo() starts the move, and again when the target changed during the move
	IF fbFollower.bStartMove THEN
		fbAxis.MoveTo();
	END_IF
	bMoveAxis := fbFollower.bMoving;
END_IF



fbAxis(
	enable 			:= bEnable,
	Reset 			:= bReset,
	HomingMode 		:= MC_ForceCalibration,
	Position 		:= fPosition, 
	Velocity 		:= fVelocity,
	Enable_Positive := TRUE,//NOT axisRef.Status.SoftLimitMaxExceeded,
	Enable_Negative := TRUE,// NOT axisRef.Status.SoftLimitMinExceeded,
	Jog_Forward 	:= bMovePos,
	Jog_Backwards 	:= bMoveNeg,
	isModuloAxis 	:= FALSE,
	ActualPosition 	=> fActualPosition,
	Error 			=> bError,
	ErrorID 		=> nErrorID,
	AxisRef 		:= axisRef);
	
IF bReset OR bError THEN
	bMoveAxis := FALSE;
END_IF

IF fbAxis.HomeDone OR bReset OR bError THEN
	bHomeAxis := FALSE;
END_IF
	
IF fbAxis.ResetDone THEN
	bReset := FALSE;
END_IF

IF fbAxis.StopDone THEN
	bStopAxis := FALSE;
END_IF


bReady := fbAxis.Ready;

fbreadParameter(	
	Axis 			:= axisRef, 
	Enable 			:= fbAxis.InMotion, 
	ParameterNumber := MC_AxisParameter.AxisRemainingTimeToGo, 
	ReadMode 		:= E_ReadMode.READMODE_CYCLIC);
				
IF fbreadParameter.Valid THEN
	fSlewtime := fbreadParameter.Value;
END_IF

HandleEvents();

// The focus has no reference switch (#22) and needs none: its encoder is absolute (the NC axis has
// ReferenceSystem ABSOLUTE and an Offset in the tsproj, the drive reports a multi-turn position), so the position
// survives an activation (test T16, 2026-10-13). Homing only sets the calibrated flag: MC_ForceCalibration ignores
// the reference position it is given and never changes the axis position. The zero point of the focus is the NC
// encoder Offset in the tsproj, not anything in the PLC. The stored position of #20 (fLastPosition) was passed
// here but never applied; #44.
METHOD _StartHoming : BOOL
fbAxis.Home(fReference := fActualPosition);		// ignored by MC_ForceCalibration
_StartHoming := TRUE;
END_METHOD

// Stop a running focus move (MC_Stop) and hold the position reached: the target becomes the actual position at
// StopDone, so the automatic positioning does not restart the move. A new Position afterwards moves again.
// Returns TRUE when an MC_Stop was requested. MONETcommon#122.
METHOD Stop : BOOL
fbFollower.Stop();
fbAxis.CancelMove();
IF fbAxis.Ready AND NOT fbAxis.StandStill THEN
	Stop := fbAxis.Stop();
	bHoldOnStop := TRUE;
ELSIF fbAxis.Calibrated THEN
	fPosition := fActualPosition;
END_IF
END_METHOD

PROPERTY PUBLIC MinPosition : LREAL
GET
MinPosition := fMinPosition;
END_GET
END_PROPERTY

PROPERTY PUBLIC MaxPosition : LREAL
GET
MaxPosition := fMaxPosition;
END_GET
END_PROPERTY

METHOD PRIVATE HandleEvents : BOOL
VAR_INPUT
END_VAR
axisEvent(	
	Trigger 		:= fbAxis.Error, 
	Level 			:= ADSLOG_MSGTYPE_ERROR,
	FormatString	:= 'Focus Axis Error: %S',
	OnMessage 		:= NCError_TO_STRING(ErrorID),
	OffMEssage 		:= 'OK',
	OffLevel 		:= ADSLOG_MSGTYPE_HINT,
	comm 			:= fbComm);

CalibrationEvent(
	Trigger 		:=	bCalibrated,
	Level 			:=	ADSLOG_MSGTYPE_HINT,
	OnMessage 		:= 'Focus Axis is calibrated.',
	comm 			:= fbComm);
END_METHOD

END_FUNCTION_BLOCK

// ---- POUs/FB_AxisControl.TcPOU
FUNCTION_BLOCK ABSTRACT FB_AxisControl EXTENDS FB_BaseAxis IMPLEMENTS I_Axis
VAR_INPUT
	bMoveAxis				: BOOL;		// Move axis to given position
	bTracking				: BOOL;		// enable tracking
	bStopAxis				: BOOL;		// stop the Axis
END_VAR
VAR_OUTPUT
END_VAR
VAR
	fSlewTime				: LREAL;	// time to reach target position
	fbAxisCalibration		:	MC_SetPosition;
	axisEvent				:	FB_EventLog;
	diagnosticEvent			:	FB_EventLog;
	
	bDiagnosticError		: BOOL;
	
	fbReadParameter			: MC_ReadParameter;
	bGetLastPosition		: BOOL := TRUE;
	
	calibrationEvent		: FB_Eventlog;
END_VAR
VAR PERSISTENT
	// UNUSED since #44: the focus used to store its position here, but the stored position was never applied (the
	// homing mode ignores it) and the focus encoder is absolute. Kept declared because removing a PERSISTENT variable
	// changes the persistent data layout; remove it together with the next layout change.
	fLastPosition			: LREAL := -1.0;
END_VAR

PROPERTY MoveAxis : BOOL
GET
MoveAxis := bMoveAxis;
END_GET
SET
// FALSE -> TRUE starts a move to fPosition (fbAxis.MoveTo(), BROTLib #63); FALSE drops a move that has not started.
// bMoveAxis stays the level the telescope sees; the axis block clears it on MoveDone.
IF MoveAxis AND NOT bMoveAxis THEN
	fbAxis.MoveTo();
ELSIF NOT MoveAxis THEN
	fbAxis.CancelMove();
END_IF
bMoveAxis := MoveAxis;
END_SET
END_PROPERTY

PROPERTY MoveDone : BOOL
GET
MoveDone := fbAxis.MoveDone;
END_GET
END_PROPERTY

PROPERTY SlewTime : LREAL
GET
SlewTime := fSlewTime;
END_GET
END_PROPERTY

PROPERTY StopAxis : BOOL
GET
StopAxis := bStopAxis;
END_GET
SET
// FALSE -> TRUE stops the axis (fbAxis.Stop(), BROTLib #63); the axis block clears bStopAxis on StopDone.
IF StopAxis AND NOT bStopAxis THEN
	fbAxis.Stop();
END_IF
bStopAxis := StopAxis;
END_SET
END_PROPERTY

PROPERTY Tracking : BOOL
GET
Tracking := bTracking;
END_GET
SET
bTracking := Tracking;
END_SET
END_PROPERTY

END_FUNCTION_BLOCK

// ---- POUs/Functions/NCError_TO_STRING.TcPOU
FUNCTION NCError_TO_STRING : STRING(255)
VAR_INPUT
	// NC Error ID
	ErrorID:	UDINT;
END_VAR
VAR
END_VAR

NCError_TO_STRING := '';

CASE ErrorID OF
	16#D012:	NCError_TO_STRING := 'Control and power section ready (no error)';
	16#D013:	NCError_TO_STRING := 'Axis in operation (no error)';
	16#4220:	NCError_TO_STRING := 'Group not ready / group not ready for new task';
	16#4253:	NCError_TO_STRING := 'Reference cam became free too soon';
	16#4257:	NCError_TO_STRING := 'Function not allowed';
	16#4260:	NCError_TO_STRING := 'Controller enable';
	16#42EF:	NCError_TO_STRING := 'Axis is locked for motion commands because a stop command is still active';
	16#4466:	NCError_TO_STRING := 'Invalid IO data FOR more than n subsequent NC cycles (encoder)';
	16#4550: 	NCError_TO_STRING := 'Following error monitoring (position)';
	16#4650:	NCError_TO_STRING := 'Drive hardware not ready to operate';
	16#4B07:	NCError_TO_STRING := 'Timeout axis function block';
	16#4B09:	NCError_TO_STRING := 'Axis is not ready';
	16#4B0A:	NCError_TO_STRING := 'Error during referencing';
	16#ECD0:	NCError_TO_STRING := 'Positive limit switch warning.';				
	16#ED43:	NCError_TO_STRING := 'Under-voltage - DC link.';				
	16#F324:	NCError_TO_STRING := 'Excessive position command value deviation';				
	16#F601:	NCError_TO_STRING := 'Calibrate commutation offset error.';				

ELSE
	NCError_TO_STRING := DWORD_TO_HEXSTR(ErrorID, 4, FALSE);
END_CASE

END_FUNCTION

// ---- POUs/FB_HourAngleControl.TcPOU
FUNCTION_BLOCK FB_HourAngleControl EXTENDS FB_AxisControl
VAR_INPUT
	bReleaseHold : BOOL;		// #159: a new power-on was accepted, release the hold (one scan, set by FB_TelescopeControl.Init)
	bStopSweep : BOOL;		// #198: a stop arrived in the calibration sweep (one scan, set by FB_TelescopeControl): hold the homing request
	fMinPosition : LREAL := -180.0;
	fMaxPosition : LREAL := 180.0;
END_VAR
VAR_OUTPUT
	bSweepActive : BOOL;		// #198: the calibration sweep is requested or running (a pause between two homing steps reports StandStill)
END_VAR
VAR
	bAxisError	: BOOL;
	bLatchHomeError	: BOOL;
	nAxisErrorID : UDINT;
	nLatchHomeErrorID: UDINT;
	bLatchHomeErrorHeld	: BOOL;		// #69: the homing error, held until the axis reset
	nLatchHomeErrorIDHeld : UDINT;
	fbLatchHome : FB_LatchHome;
	fbHomeHold : FB_HomeHold;		// #113: no homing request after a stop of the axis
	tonReady : TON;					// #155: the NC axis takes some time after Ready before a command reaches it
	bResetForAbort : BOOL;		// #113: the reset was asked for by FB_LatchHome to end a homing, it must not release the hold
	omega 	: LREAL := 360.0 / 86164.099 * (PI/180.0); //sidereal velocity
END_VAR

// limit to sane positions
fPosition := LIMIT(fMinPosition, fPosition, fMaxPosition);


// #113: a stop during the calibration sweep must not be followed by a new homing request (bHomeAxis was set again every
// scan while the axis is enabled and uncalibrated, so FB_LatchHome went on commanding the NC while MC_Stop held the lock)
// #113: FB_LatchHome asks for a reset when MC_AbortHoming cannot end a running step. That reset must not release the hold
// (the sweep would start again); the hold ends with the disable that FB_SweepStop does after the stop.
IF fbLatchHome.ResetRequest THEN
	bReset := TRUE;
	bResetForAbort := TRUE;
END_IF
IF NOT bEnable THEN
	bResetForAbort := FALSE;
END_IF
fbHomeHold(bEnable := bEnable, bCalibrated := fbAxis.Calibrated, bHoming := bHomeAxis, bStopAxis := bStopAxis, bReset := bReset AND NOT bResetForAbort, bRelease := bReleaseHold, bStopSweep := bStopSweep);
bReleaseHold := FALSE;
bStopSweep := FALSE;

// #155: not before the NC axis is enabled, and not right after Ready either: the first reference step started 5 to 40 ms
// after Ready still aborts about 80 ms later, and the abort and the re-arm can overlap (4B66). Ready for 0.5 s.
tonReady(IN := bEnable AND fbAxis.Ready, PT := T#500MS);
IF tonReady.Q AND NOT fbAxis.Calibrated AND NOT fbHomeHold.bHold THEN
	bHomeAxis := TRUE;
END_IF

// #155: the request used to survive a disable. After the next enable it was already TRUE, so FB_LatchHome saw no rising
// edge and the sweep never started.
IF fbAxis.Calibrated OR fbHomeHold.bHold OR NOT bEnable THEN
	bHomeAxis := FALSE;
END_IF

IF bHomeAxis THEN
	fPosition := fPosition;
END_IF

fbAxis(
	enable 			:= bEnable,
	Reset 			:= bReset,
	Tracking 		:= bTracking,
	HomingMode 		:= MC_ForceCalibration,
	Position 		:= fPosition, 
	Velocity 		:= fVelocity,
	TrackVelocityRef	:= omega,
	TrackDirectionRef:=0,
	Enable_Positive := NOT axisRef.Status.SoftLimitMaxExceeded,
	Enable_Negative := NOT axisRef.Status.SoftLimitMinExceeded,
	Jog_Forward 	:= bMovePos,
	Jog_Backwards 	:= bMoveNeg,
	ActualPosition 	=> fActualPosition,
	Error 			=> bAxisError,
	ErrorID 		=> nAxisErrorID,
	AxisRef 		:= axisRef);

// #100: follow the NC in both directions. The flag used to be set only while the axis was calibrated, so it stayed
// TRUE after the NC dropped Homed and the power-on and bHomed trusted it.
bCalibrated := fbAxis.Calibrated;

fbLatchHome(
	Axis				:= AxisRef,
	Execute				:= bHomeAxis,
	Reset				:= bReset,	// #155
	StopActive			:= bStopAxis OR ((axisRef.NcToPlc.StateDWord AND 16#20000000) <> 0),	// #113
	Direction 			:= MC_Home_Direction.mcPositiveDirection,
	Velocity 			:= 1.0,
	Acceleration		:= 3.6,
	Deceleration		:= 3.6,
	Jerk				:= 3.6,
	RefPosition			:= 1.56-0.04019852332911753,
	RefDistance			:= 5.21,
	TimeLimit 			:= T#1M,
	DistanceLimit 		:= 6,
	TravelLimit			:= 21,	// #165: 3 steps of 6 deg and the 2 deg jog, plus a margin
	Error 				=> bLatchHomeError,
	ErrorID 			=> nLatchHomeErrorID);
	

// #198
bSweepActive := bHomeAxis OR fbLatchHome.Busy;

// #69: FB_LatchHome clears its error as soon as Execute falls, and Execute falls on bError, so the error lasted
// one scan: the power-on was aborted, bError was FALSE again and no reset could fire. Hold it until the axis reset.
IF bReset THEN
	bLatchHomeErrorHeld := FALSE;
	nLatchHomeErrorIDHeld := 0;
END_IF
IF bLatchHomeError THEN
	bLatchHomeErrorHeld := TRUE;
	nLatchHomeErrorIDHeld := nLatchHomeErrorID;
END_IF

bError := bLatchHomeErrorHeld OR bAxisError;

// nErrorID is the current error: it used to keep stale values, so healthy axes were reset on every reset pass
IF bAxisError THEN
	nErrorID := nAxisErrorID;
ELSIF bLatchHomeErrorHeld THEN
	nErrorID := nLatchHomeErrorIDHeld;
ELSE
	nErrorID := 0;
END_IF
	
IF fbAxis.MoveDone OR bReset OR bError THEN
	bMoveAxis := FALSE;
END_IF

IF (fbAxis.HomeDone AND fbLatchHome.Done) OR bReset OR bError THEN
	bHomeAxis := FALSE;
END_IF
	
IF fbAxis.ResetDone THEN
	bReset := FALSE;
END_IF

// #159: bStopAxis was cleared only on StopDone. A stop of an axis that is disabled or standing still gives none, so
// it stayed TRUE and held every following sweep until a Reset Cold.
IF fbAxis.StopDone OR NOT bEnable OR bReset THEN
	bStopAxis := FALSE;
END_IF


bReady := fbAxis.Ready;

fbReadParameter(	
	Axis 			:= axisRef, 
	Enable 			:= fbAxis.InMotion, 
	ParameterNumber := MC_AxisParameter.AxisRemainingTimeToGo, 
	ReadMode 		:= E_ReadMode.READMODE_CYCLIC);
				
IF fbReadParameter.Valid THEN
	fSlewtime := fbReadParameter.Value;
END_IF


axisEvent(	
	Trigger 		:= bError, 
	Level 			:= ADSLOG_MSGTYPE_ERROR,
	FormatString	:= 'Hour Angle Axis Error: %s',
	OnMessage 		:= NCError_TO_STRING(nErrorID),
	OffMEssage 		:= 'OK',
	OffLevel 		:= ADSLOG_MSGTYPE_HINT,
	Comm			:= fbComm);
	

CalibrationEvent(	
	Trigger 		:= bCalibrated, 
	Level 			:= ADSLOG_MSGTYPE_HINT,
	OnMessage 		:= 'Hour Angle Axis is calibrated.',
	Comm			:= fbComm);

// Homing goes through FB_LatchHome and MC_SetPosition on bHomeAxis (the level), not through fbAxis.Home(), so this
// is empty (abstract in BROTLib's FB_BaseAxis, BROTLib #62).
METHOD _StartHoming : BOOL
_StartHoming := TRUE;
END_METHOD

END_FUNCTION_BLOCK

// ---- POUs/FB_LatchHome.TcPOU
FUNCTION_BLOCK FB_LatchHome

VAR_IN_OUT
	Axis						: AXIS_REF;
END_VAR
VAR_INPUT
	Execute					: BOOL;										(* B *)
	StopActive				: BOOL;										(* #113: the axis is being stopped (stop requested or MC_Stop lock): abort the sequence *)
	Reset					: BOOL;										(* #155: leave the abort state at once, whatever MC_AbortHoming does *)

	(* static parameters *)
	Direction					: MC_Home_Direction;						(* E *)
	

	Velocity					: LREAL;									(* E *)
	Acceleration				: LREAL;									(* V *)	(* Beckhoff proprietary input *)
	Deceleration				: LREAL;									(* V *)	(* Beckhoff proprietary input *)
	Jerk						: LREAL;									(* V *)	(* Beckhoff proprietary input *)
	
	MoveIsCountDirection		: BOOL := TRUE;								(* If not specified : TRUE *)

	RefPosition					: LREAL;									(* Position (physical) of first marker of RefDistance in travel direction [deg]*)
	RefDistance					: LREAL; 									(* Reference distance to calibrate Latch distances to physical coords. ( >5.00 deg!!!)*)
	(* maximum time for one ref search process *)
	TimeLimit					: TIME;										(* E *)

	(* maximum travel distance for on calibration step (should be 6) *)
	DistanceLimit				: LREAL;									(* E *)
	(* #165: maximum distance of the axis from where the sequence started, over all segments and restarts (0 = off). The
	   limit per step does not bound the sequence: 3 steps out, a jog and 3 back, and an abort restarts it. *)
	TravelLimit				: LREAL;
	
	(* Set bipolar torque limit to this value to avoid mechanical damadges [%] *)
	TorqueLimit					: LREAL;								(* E *)

	BufferMode					: MC_BufferMode;							(* E *)
	Options						: ST_Home_Options4;
END_VAR
VAR_OUTPUT
	Done						: BOOL;										(* B *)
	Busy						: BOOL;										(* E *)
	Active						: BOOL;										(* E *)
	CommandAborted				: BOOL;										(* E *)
	Error						: BOOL;										(* B *)
	ErrorID						: UDINT;									(* E *)
	ResetRequest				: BOOL;										(* #113: the axis is to be reset to end a homing that MC_AbortHoming cannot abort *)
END_VAR
VAR	
	RefSignal					: MC_Ref_Signal_Ref;
	ReadApplicationRequest		: MC_ReadApplicationRequest;
	ApplicationRequest			: ST_NcApplicationRequest;

	Parameter					: MC_HomingParameter;

	Axis_Status:	MC_ReadStatus;
	Axis_Power:		MC_Power;
	
	bEnable						: BOOL;
	bReady						: BOOL;
	bCalibrated					: BOOL;

	Request						: BOOL;		(* application request bit [0/1] *)
	RequestType					: UINT;		(* application request TYPE/ID *)

	StepReferencePulseDetection			: MC_StepReferencePulseDetection;
	MoveAxis					: MC_Jog;

	SetPos						: MC_SetPosition;
	
	StepFinishHoming			: MC_FinishHoming;
	StepAbortHoming				: MC_AbortHoming;
	
	(* Need three Ref positions for absolut calibration *)
	(* One way *)
	RecordedPositions_to		: ARRAY [0..2] OF LREAL;
	(* Going back for checking*)
	RecordedPositions_back		: ARRAY [0..2] OF LREAL;
	
	RecordedDistances_to		: ARRAY [0..1] OF LREAL;
	RecordedDistances_back		: ARRAY [0..1] OF LREAL;
	
	PostionReset				: ARRAY [0..2] OF LREAL := [0,0,0];
	DistanceReset				: ARRAY [0..1] OF LREAL := [0,0];
	
	PositionOffset				: LREAL;
	iErrorId					: UDINT;
	iCommandAborted				: BOOL;
	
	nState						: INT;
	nAbortFrom					: INT;									(* #113: state in which the sequence was aborted *)
	bRearm						: BOOL;									(* #155: re-arm the start once the abort has settled *)
	fbRearmDelay				: TON;
	bTakeStart					: BOOL;
	fbStepDrain					: FB_StepDrain;							(* #113: drain of a stale step block before a start *)
	bStepBusy					: BOOL;									(* #113: a step block is still running its NC command *)
	nSearch						: INT;
	fStartPos					: LREAL;								(* #165: axis position before the sequence started, sampled while Execute is FALSE *)
	bTravelExceeded			: BOOL;									(* #165 *)

	fbStartReq					: FB_StartRequest;						(* #155: start request, kept until state 0 can take it *)
	fbReady						: R_TRIG;
	fbTimeOut					: TON;
	fbLockWait					: TON;									(* #113: longest wait for the MC_Stop lock before MC_AbortHoming *)
	fbAbortTimeout				: TON;									(* #155: longest time in the abort state, it has no other exit *)
END_VAR
VAR CONSTANT
	ERR_ABORT_TIMEOUT			: UDINT := 16#4F000001;					(* #155: the abort did not finish in time *)
	ERR_STEP_STUCK				: UDINT := 16#4F000002;					(* #113: a step block does not leave Busy, no start possible *)
	ERR_TRAVEL_LIMIT			: UDINT := 16#4F000003;					(* #165: the search left the allowed range without finding the marks *)
END_VAR

// #155: the rising edge of Execute is only taken in state 0. One that arrives while the sequence is still aborting would
// be lost and the axis would never start, so remember it until state 0 is reached (and drop it with Execute).
fbStartReq(Execute := Execute);

RefSignal.TouchProbe := E_TouchProbe.TouchProbe1;

// #113: nothing else stops this sequence (a step block ignores a falling Execute, and the state machine reads Execute
// only in state 0). A stop of the axis, or Execute going away, aborts it: release the step blocks and go to the abort
// state, which waits for the MC_Stop lock to clear.
// #165: the sample is not taken after a start, so a restart after an abort (Execute stays TRUE) keeps the first start
IF nState = 0 AND NOT Execute THEN
	fStartPos := Axis.NcToPlc.ActPos;
END_IF
bTravelExceeded := TravelLimit > 0 AND nState >= 1 AND nState <= 3 AND ABS(Axis.NcToPlc.ActPos - fStartPos) > TravelLimit;
IF nState >= 1 AND nState <= 6 AND (NOT Execute OR StopActive OR bTravelExceeded) THEN
	nAbortFrom := nState;
	// #113 mode 2: the running reference step keeps its Execute until the abort is over
	IF GVL_Homing.nAbortMode <> 2 THEN
		StepReferencePulseDetection(
			Execute					:= FALSE,
			Parameter				:= Parameter,
			Axis					:= Axis);
	END_IF
	MoveAxis(
		Axis					:= Axis,
		JogForward				:= FALSE,
		JogBackwards			:= FALSE);
	SetPos(
		Execute					:= FALSE,
		Axis					:= Axis);
	StepFinishHoming(
		Execute					:= FALSE,
		Parameter				:= Parameter,
		Axis					:= Axis);
	iErrorId := 0;
	IF bTravelExceeded THEN
		iErrorId := ERR_TRAVEL_LIMIT;
	END_IF
	nState := 20;
END_IF
fbLockWait(IN := nState = 20 AND StopActive AND NOT StepAbortHoming.Busy, PT := T#5S);
fbAbortTimeout(IN := nState = 20, PT := T#10S);
// #155: not in the scan in which the abort ended: the NC has to settle, a start at once overlapped it (4B66)
fbRearmDelay(IN := bRearm AND nState = 0 AND Execute, PT := T#300MS);
IF fbRearmDelay.Q THEN
	bRearm := FALSE;
	fbStartReq.Rearm();
ELSIF NOT Execute THEN
	bRearm := FALSE;
END_IF
ResetRequest := FALSE;
bStepBusy := StepReferencePulseDetection.Busy OR MoveAxis.Busy OR SetPos.Busy OR StepFinishHoming.Busy;
// #113: a stop leaves the reference step Busy (it ignores the falling Execute), and the reset of the axis ends its NC command
// without the block ever being called again. At the next start it then reported the old command as finished, the sequence
// went to the abort state and the abort overlapped the new MC_Home (4B66). In state 0 call a Busy block with FALSE until it
// drops Busy, and take no start before.
fbStepDrain(bIdle := nState = 0, bStepBusy := bStepBusy, bStartPending := fbStartReq.Pending);
IF fbStepDrain.bStuck THEN
	fbStartReq.Take();
	Error := TRUE;
	ErrorID := ERR_STEP_STUCK;
END_IF

CASE nState OF
	0 :	(* init *)
		IF fbStepDrain.bDrain THEN
			StepReferencePulseDetection(
				Execute					:= FALSE,
				Parameter				:= Parameter,
				Axis					:= Axis);
			MoveAxis(
				Axis					:= Axis,
				JogForward				:= FALSE,
				JogBackwards			:= FALSE);
			SetPos(
				Execute					:= FALSE,
				Axis					:= Axis);
			StepFinishHoming(
				Execute					:= FALSE,
				Parameter				:= Parameter,
				Axis					:= Axis);
		END_IF
		// #113 mode 2: release the reference step that was kept running during the abort
		IF GVL_Homing.nAbortMode = 2 THEN
			StepReferencePulseDetection(
				Execute					:= FALSE,
				Parameter				:= Parameter,
				Axis					:= Axis);
		END_IF
		IF NOT Execute THEN
			(* reset at falling edge of Execute *)
			Busy 			:= FALSE;
			Done			:= FALSE;
			CommandAborted 	:= FALSE;
			Error 			:= FALSE;
			ErrorID 		:= 0;
			iErrorID 		:= 0;
			
			bEnable			:= FALSE;
			
			nSearch 		:= 0;
			
			//Reset Arrays to zeros
			RecordedPositions_to	:= PostionReset;
			RecordedPositions_back	:= PostionReset;
			RecordedDistances_to	:= DistanceReset;
			RecordedDistances_back	:= DistanceReset;
		END_IF
 	
		IF fbStepDrain.bMayTake THEN
			bTakeStart := fbStartReq.Take();
		ELSE
			bTakeStart := FALSE;
		END_IF
	  	IF bTakeStart THEN
			(* initialize output values *)
	  		Busy 				:= TRUE;

			IF BufferMode <> 0 THEN
				Busy := FALSE;
				Error := TRUE;
				ErrorID := MC_ERROR_BUFFERMODE_NOT_SUPPORTED;

				nState := 0;
			ELSE
				(* For axis with non Beckhoff components -> needs to be true (don't get why)*)
				Options.DisableDriveAccess := TRUE;
				nSearch:=0;
				nState := nState + 1; 
			END_IF
		END_IF
	1: (* Search one Block *)
		StepReferencePulseDetection(
			Execute 			:= TRUE,
			Direction 			:= Direction,
			ReferenceSignal 	:= RefSignal,
			Velocity 			:= Velocity,
			Acceleration 		:= Acceleration,
			Deceleration 		:= Deceleration,
			Jerk				:= Jerk,
			TimeLimit 			:= TimeLimit,
			TorqueLimit			:= TorqueLimit,
			DistanceLimit 		:= DistanceLimit,
			Axis				:= Axis,
			Parameter			:= Parameter,
			BufferMode			:= BufferMode, 
			Options				:= Options, 
			RecordedPosition	=> RecordedPositions_to[nSearch]);
			
		IF NOT StepReferencePulseDetection.Busy AND StepReferencePulseDetection.Done THEN
			StepReferencePulseDetection(	
				Execute					:= FALSE, 
				Parameter				:= Parameter,
				Axis					:= Axis);
			nSearch := nSearch +1;
			IF nSearch >2 THEN
				nState := nState + 1;
			END_IF

			
		ELSIF NOT StepReferencePulseDetection.Busy AND (StepReferencePulseDetection.Error OR StepReferencePulseDetection.CommandAborted) THEN
			iErrorID := StepReferencePulseDetection.ErrorID; 					(* functional/calibration error *) (* HKP *)
			
			StepReferencePulseDetection(	
				Execute					:= FALSE, 
				Parameter				:= Parameter,
				Axis					:= Axis);

			nState 	:= 20;
		END_IF
	2:	(* Jog 2 degrees *)
		nSearch := 0;
		IF Direction = MC_Home_Direction.mcPositiveDirection THEN
			MoveAxis.JogForward := TRUE;
		ELSIF Direction = MC_Home_Direction.mcNegativeDirection THEN
			MoveAxis.JogBackwards := TRUE;
		ELSE
			iErrorID := 1;
			nState := 20;
		END_IF
		MoveAxis(
			Axis				:= Axis,	
			Mode 				:= E_JogMode.MC_JOGMODE_INCHING,
			JogForward			:=,
			JogBackwards		:=,
			Position			:= 2,
			Velocity 			:= Velocity,
			Acceleration 		:= Acceleration,
			Deceleration 		:= Deceleration,
			Jerk				:= Jerk);
		IF NOT MoveAxis.Busy AND MoveAxis.Done THEN
			MoveAxis(	
				Axis				:= Axis,
				JogForward			:= FALSE,
				JogBackwards		:= FALSE);
			nState := nState + 1;

			
		ELSIF NOT MoveAxis.Busy AND (MoveAxis.Error OR MoveAxis.CommandAborted) THEN
			iErrorID := MoveAxis.ErrorID; 					(* functional/calibration error *) (* HKP *)
			
			MoveAxis(	
				Axis				:= Axis,
				JogForward			:= FALSE,
				JogBackwards		:= FALSE);

			nState 	:= 20;
		END_IF
		
	3:	(* Search two Block *)
		// Change Direction to move backwards
		IF Direction = MC_Home_Direction.mcPositiveDirection THEN
			StepReferencePulseDetection.Direction := MC_Home_Direction.mcNegativeDirection;
		ELSIF Direction = MC_Home_Direction.mcNegativeDirection THEN
			StepReferencePulseDetection.Direction := MC_Home_Direction.mcPositiveDirection;
		ELSE
			iErrorID := 1;
			nState := 20;
		END_IF
		StepReferencePulseDetection(
			Execute 			:= TRUE,
			Direction 			:=,
			ReferenceSignal 	:= RefSignal,
			Velocity 			:= Velocity,
			Acceleration 		:= Acceleration,
			Deceleration 		:= Deceleration,
			Jerk				:= Jerk,
			TimeLimit 			:= TimeLimit,
			TorqueLimit			:= TorqueLimit,
			DistanceLimit 		:= DistanceLimit,
			Axis				:= Axis,
			Parameter			:= Parameter,
			BufferMode			:= BufferMode, 
			Options				:= Options, 
			RecordedPosition	=> RecordedPositions_back[nSearch]);
			
		IF NOT StepReferencePulseDetection.Busy AND StepReferencePulseDetection.Done THEN
			StepReferencePulseDetection(	
				Execute					:= FALSE, 
				Parameter				:= Parameter,
				Axis					:= Axis);
			nSearch := nSearch +1;
			IF nSearch >2 THEN
				nState := nState + 1;
			END_IF

			
		ELSIF NOT StepReferencePulseDetection.Busy AND (StepReferencePulseDetection.Error OR StepReferencePulseDetection.CommandAborted) THEN
			iErrorID := StepReferencePulseDetection.ErrorID; 					(* functional/calibration error *) (* HKP *)
			
			StepReferencePulseDetection(	
				Execute					:= FALSE, 
				Parameter				:= Parameter,
				Axis					:= Axis);

			nState 	:= 20;
		END_IF
	4: (* Calculate Distances*)
		nSearch:=0;
		FOR nSearch:=0 TO 1 BY 1 DO
			RecordedDistances_to[nSearch] := F_RoundLREAL(ABS(RecordedPositions_to[nSearch] - RecordedPositions_to[nSearch+1]), 2);
			RecordedDistances_back[nSearch] := F_RoundLREAL(ABS(RecordedPositions_back[nSearch] - RecordedPositions_back[nSearch+1]), 2);
		END_FOR
		IF RecordedDistances_to[0] = RecordedDistances_back[1] AND RecordedDistances_to[1] = RecordedDistances_back[0] THEN
			nState := nState +1;
		ELSE
			(*if distances changed -> something is truely wrong*)
			iErrorID:=1;
			nState := 20;
		END_IF
	
	5: (* look up distance gaps and then set position and reference flag *)
		SetPos.Options.ClearPositionLag := TRUE;
		
		IF RefDistance > 5.0 THEN
			IF MoveIsCountDirection THEN
				IF RecordedDistances_to[0] > 5 THEN
					PositionOffset := (RecordedDistances_to[0] - RefDistance)*1000 + RefPosition - RecordedPositions_to[0];
				ELSE
					PositionOffset := (RecordedDistances_to[1] - RefDistance)*1000 + RefPosition - RecordedPositions_to[1];
				END_IF
			ELSE
				IF RecordedDistances_to[0] > 5 THEN
					PositionOffset := -(RecordedDistances_to[0] - RefDistance)*1000 + RefPosition - RecordedPositions_to[0];
				ELSE
					PositionOffset := -(RecordedDistances_to[1] - RefDistance)*1000 + RefPosition - RecordedPositions_to[1];
				END_IF
			END_IF
		ELSE
			iErrorID := 1;
			nState := 20;
		END_IF
		
		
		SetPos(
			Axis				:= Axis, 
			Execute				:= TRUE, 
			Position			:= PositionOffset, 
			Mode				:= TRUE, // relative postion change
			Options				:= );

		IF NOT SetPos.Busy AND SetPos.Done THEN
			SetPos(	
				Execute					:= FALSE, 
				Axis					:= Axis);

			nState := nState + 1;
		ELSIF NOT SetPos.Busy AND SetPos.Error THEN
			iErrorID := SetPos.ErrorID; (* functional/calibration error *)

			SetPos(	
				Execute					:= FALSE, 
				Axis					:= Axis);

			nState 	:= 20;
		END_IF
	
	6:
		StepFinishHoming.Options.DisableDriveAccess := Options.DisableDriveAccess;
		
		StepFinishHoming(	
			Execute				:= TRUE, 
			Distance			:= , 
			Velocity			:= Velocity, 
			Acceleration		:= Acceleration, 
			Deceleration		:= Acceleration, 
			Jerk				:= Jerk, 
			BufferMode			:= BufferMode, 
			Options				:= , 
			Axis				:= Axis, 
			Parameter			:= Parameter); 

		IF NOT StepFinishHoming.Busy AND StepFinishHoming.Done THEN
			Busy 				:= FALSE;
			Done	 			:= TRUE;

			StepFinishHoming(	
				Execute					:= FALSE, 
				Parameter				:= Parameter,
				Axis					:= Axis);

			nState := 0; 
		ELSIF NOT StepFinishHoming.Busy AND (StepFinishHoming.Error OR StepFinishHoming.CommandAborted) THEN
			iErrorID 		:= StepFinishHoming.ErrorID;

			StepFinishHoming(
				Execute					:= FALSE, 
				Parameter				:= Parameter,
				Axis					:= Axis);

			nState := 20;
		END_IF

	20:	(*Abort Homing*)
		// #155: no other exit: a reset or the timeout leaves the state even if MC_AbortHoming never reports back
		IF Reset OR fbAbortTimeout.Q THEN
			StepAbortHoming(
				Axis				:= Axis,
				Parameter			:= Parameter,
				Execute				:= FALSE,
				Options				:= );
			Busy := FALSE;
			IF Reset THEN
				CommandAborted := TRUE;
			ELSE
				Error := TRUE;
				ErrorID := ERR_ABORT_TIMEOUT;
			END_IF
			nState := 0;
		ELSE
		// #113: MC_Stop locks the axis for motion commands until it is done (StateDWord bit 29); MC_AbortHoming sent into the
		// lock is rejected (17135) and the error disables both axes. Wait for the lock to clear, 5 s at most.
		IF NOT StopActive OR fbLockWait.Q OR StepAbortHoming.Busy THEN
			IF GVL_Homing.nAbortMode = 1 AND bStepBusy AND NOT StepAbortHoming.Busy THEN
				// #113 mode 1: MC_AbortHoming into a running step never completes (HomingBusy stays TRUE, 4F000001 after
				// 10 s), but a reset of the axis does end it. Ask for one; the Reset input then leaves this state.
				ResetRequest := TRUE;
			ELSE
			StepAbortHoming.Options.DisableDriveAccess := Options.DisableDriveAccess AND (GVL_Homing.nAbortMode <> 3);
			IF GVL_Homing.nAbortMode = 2 AND (nAbortFrom = 1 OR nAbortFrom = 3) THEN
				StepReferencePulseDetection(
					Execute					:= TRUE,
					Parameter				:= Parameter,
					Axis					:= Axis);
			END_IF

			StepAbortHoming(
				Axis				:= Axis, 
				Parameter			:= Parameter, 
				Execute				:= TRUE, 
				Options				:= ); 

			IF NOT StepAbortHoming.Busy AND StepAbortHoming.Done THEN
				Busy 				:= FALSE;
				IF iErrorId <> 0 THEN
					Error	 			:= TRUE;
					ErrorId				:= iErrorId;
				ELSE
					CommandAborted		:= TRUE;
					// #155: aborted by itself (not by a stop, a reset or Execute going away): the start is still
					// requested, so request it again. Execute stays TRUE, there is no new edge to do it.
					IF Execute AND NOT StopActive AND NOT Reset THEN
						bRearm := TRUE;
					END_IF
				END_IF
		
				StepAbortHoming(	
					Execute					:= FALSE, 
					Parameter				:= Parameter,
					Axis					:= Axis);

				nState := 0; 
			ELSIF NOT StepAbortHoming.Busy AND StepAbortHoming.Error THEN
				Busy := FALSE;
				Error := TRUE;
				ErrorID 		:= StepAbortHoming.ErrorID;

				StepAbortHoming(
					Execute					:= FALSE, 
					Parameter				:= Parameter,
					Axis					:= Axis);

				nState := 0;
			END_IF
			END_IF
		END_IF
		END_IF

END_CASE

END_FUNCTION_BLOCK

// ---- POUs/FB_StepDrain.TcPOU
// Decides what FB_LatchHome does with a step block that is still Busy while it is idle (#113). A stop leaves the reference
// step Busy and the reset of the axis ends its NC command without the block being called again; at the next start the block
// reported the old command as aborted and the abort overlapped the new MC_Home (4B66). While idle a Busy block is called with
// Execute FALSE until it drops Busy, and no start is taken before. Pure logic, tested offline in IAG50cmTests (the offline
// mocks do not run FB_LatchHome).
FUNCTION_BLOCK FB_StepDrain
VAR_INPUT
	bIdle			: BOOL;		// FB_LatchHome is in state 0
	bStepBusy		: BOOL;		// a step block still runs its NC command
	bStartPending	: BOOL;		// a start request waits to be taken
	PT				: TIME := T#2S;	// longest wait for the step block to leave Busy while a start is pending
END_VAR
VAR_OUTPUT
	bDrain			: BOOL;		// call the step blocks with Execute FALSE
	bMayTake		: BOOL;		// a pending start may be taken
	bStuck			: BOOL;		// the step block did not leave Busy in time: give up the start
END_VAR
VAR
	fbStuck			: TON;
END_VAR

bDrain := bIdle AND bStepBusy;
bMayTake := bIdle AND NOT bStepBusy;
fbStuck(IN := bDrain AND bStartPending, PT := PT);
bStuck := fbStuck.Q;

END_FUNCTION_BLOCK

// ---- POUs/FB_StartRequest.TcPOU
// A start request that is kept until it is taken (#155). FB_LatchHome read the rising edge of Execute only in its idle
// state, so an edge that arrived while the sequence was still aborting was lost: Execute stayed TRUE, no new edge came,
// the axis never started its calibration and the power-on waited in stage 40 for good. The request is dropped when
// Execute falls, and taking it does not restart anything while Execute stays TRUE. Pure logic, tested offline in IAG50cmTests.
FUNCTION_BLOCK FB_StartRequest
VAR_INPUT
	Execute		: BOOL;
END_VAR
VAR_OUTPUT
	Pending		: BOOL;		// a start was requested and not taken yet
END_VAR
VAR
	fbEdge		: R_TRIG;
END_VAR

fbEdge(CLK := Execute);
Pending := (Pending OR fbEdge.Q) AND Execute;

METHOD Rearm
// a start that ended without a result while Execute is still TRUE: there is no new edge, ask again
Pending := Execute;
END_METHOD

METHOD Take : BOOL
Take := Pending;
Pending := FALSE;
END_METHOD

END_FUNCTION_BLOCK

// ---- POUs/Functions/F_RoundLREAL.TcPOU
FUNCTION F_RoundLREAL : LREAL
VAR_INPUT
  rInput : LREAL;
  iDecimalPlaces : INT;
END_VAR
VAR
  rOutput : LREAL;
  rLeftPart : LREAL;
END_VAR

(*
Source: https://medium.com/@hristo.iliev.ganchev/how-to-round-a-real-lreal-in-twincat-d551172555f3
Date: 2023–29–08
Author: Hristo Ganchev (https://github.com/hganchev)

Adapted from REAL to LREAL
*)


rOutput := rInput * EXPT(10,iDecimalPlaces);
rLeftPart := rOutput - LTRUNC(rOutput);

IF rLeftPart >= 0.5 THEN
  rOutput := rOutput + 1;
ELSIF rLeftPart <= -0.5 THEN
  rOutput := rOutput - 1;
ELSE
  rOutput := rOutput;
END_IF

rOutput :=  LTRUNC(rOutput) / EXPT(10,iDecimalPlaces);
F_RoundLREAL := rOutput;

END_FUNCTION

// ---- POUs/FB_HomeHold.TcPOU
// No new homing request after a stop of the axis (#113). The axis blocks used to set bHomeAxis again every scan while the
// axis is enabled and uncalibrated, so a stop in the calibration sweep did not end the sweep: FB_LatchHome went on
// commanding the NC while MC_Stop held the axis locked (error 17135, both axes disabled). A stop request while the axis
// is homing holds the request until the axis is disabled or reset. Pure logic, tested offline in IAG50cmTests.
FUNCTION_BLOCK FB_HomeHold
VAR_INPUT
	bEnable		: BOOL;		// the axis is enabled
	bCalibrated	: BOOL;
	bHoming		: BOOL;		// bHomeAxis: the calibration sweep is requested
	bStopAxis	: BOOL;		// a stop of the axis is requested (cleared on StopDone)
	bReset		: BOOL;
	bRelease	: BOOL;		// #159: a new power-on was accepted
	bStopSweep	: BOOL;		// #198: a stop arrived in the sweep (one scan): hold even if the sweep has not started yet
END_VAR
VAR_OUTPUT
	bHold		: BOOL;		// do not request homing
END_VAR

IF ((bStopAxis AND bHoming) OR bStopSweep) AND NOT bCalibrated THEN
	bHold := TRUE;
END_IF
// #159: an automatic stop (horizon, pole, calibration lost) leaves the axes enabled with the hold set, and reset=1 gives no
// bReset without an error. A new power-on releases it, but never through a stop that is still running.
IF NOT bEnable OR bReset OR (bRelease AND NOT bStopAxis AND NOT bStopSweep) THEN
	bHold := FALSE;
END_IF

END_FUNCTION_BLOCK

// ---- POUs/FB_DeclinationControl.TcPOU
FUNCTION_BLOCK FB_DeclinationControl EXTENDS FB_AxisControl
VAR_INPUT
	bReleaseHold : BOOL;		// #159: a new power-on was accepted, release the hold (one scan, set by FB_TelescopeControl.Init)
	bStopSweep : BOOL;		// #198: a stop arrived in the calibration sweep (one scan, set by FB_TelescopeControl): hold the homing request
	fMinPosition : LREAL := -50.0;
	fMaxPosition : LREAL := 180.0;
END_VAR
VAR_OUTPUT
	bSweepActive : BOOL;		// #198: the calibration sweep is requested or running (a pause between two homing steps reports StandStill)
END_VAR
VAR
	bAxisError : BOOL;
	bLatchHomeError	: BOOL;
	nAxisErrorID : UDINT;
	nLatchHomeErrorID: UDINT;
	bLatchHomeErrorHeld	: BOOL;		// #69: the homing error, held until the axis reset
	nLatchHomeErrorIDHeld : UDINT;
	fbLatchHome : FB_LatchHome;
	fbHomeHold : FB_HomeHold;		// #113: no homing request after a stop of the axis
	tonReady : TON;					// #155: the NC axis takes some time after Ready before a command reaches it
	bResetForAbort : BOOL;		// #113: the reset was asked for by FB_LatchHome to end a homing, it must not release the hold
END_VAR

// limit to sane positions
fPosition := LIMIT(fMinPosition, fPosition, fMaxPosition);


// #113: a stop during the calibration sweep must not be followed by a new homing request (bHomeAxis was set again every
// scan while the axis is enabled and uncalibrated, so FB_LatchHome went on commanding the NC while MC_Stop held the lock)
// #113: FB_LatchHome asks for a reset when MC_AbortHoming cannot end a running step. That reset must not release the hold
// (the sweep would start again); the hold ends with the disable that FB_SweepStop does after the stop.
IF fbLatchHome.ResetRequest THEN
	bReset := TRUE;
	bResetForAbort := TRUE;
END_IF
IF NOT bEnable THEN
	bResetForAbort := FALSE;
END_IF
fbHomeHold(bEnable := bEnable, bCalibrated := fbAxis.Calibrated, bHoming := bHomeAxis, bStopAxis := bStopAxis, bReset := bReset AND NOT bResetForAbort, bRelease := bReleaseHold, bStopSweep := bStopSweep);
bReleaseHold := FALSE;
bStopSweep := FALSE;

// #155: not before the NC axis is enabled, and not right after Ready either: the first reference step started 5 to 40 ms
// after Ready still aborts about 80 ms later, and the abort and the re-arm can overlap (4B66). Ready for 0.5 s.
tonReady(IN := bEnable AND fbAxis.Ready, PT := T#500MS);
IF tonReady.Q AND NOT fbAxis.Calibrated AND NOT fbHomeHold.bHold THEN
	bHomeAxis := TRUE;
END_IF

// #155: the request used to survive a disable. After the next enable it was already TRUE, so FB_LatchHome saw no rising
// edge and the sweep never started.
IF fbAxis.Calibrated OR fbHomeHold.bHold OR NOT bEnable THEN
	bHomeAxis := FALSE;
END_IF

IF bHomeAxis THEN
	fPosition := fPosition;
END_IF

fbAxis(
	enable 			:= bEnable,
	Reset 			:= bReset,
	Tracking 		:= bTracking,
	HomingMode 		:= MC_ForceCalibration,
	Position 		:= fPosition, 
	Velocity 		:= fVelocity,
	TrackVelocityRef:= 0.0,
	TrackDirectionRef:= 0,
	Enable_Positive := NOT axisRef.Status.SoftLimitMaxExceeded,
	Enable_Negative := NOT axisRef.Status.SoftLimitMinExceeded,
	Jog_Forward 	:= bMovePos,
	Jog_Backwards 	:= bMoveNeg,
	ActualPosition 	=> fActualPosition,
	Error 			=> bAxisError,
	ErrorID 		=> nAxisErrorID,		// was nErrorID: nAxisErrorID below was never written, so every Dec error read 0 (#55)
	AxisRef 		:= axisRef);
	
// #100: follow the NC in both directions. The flag used to be set only while the axis was calibrated, so it stayed
// TRUE after the NC dropped Homed and the power-on and bHomed trusted it.
bCalibrated := fbAxis.Calibrated;

fbLatchHome(
	Axis				:= AxisRef,
	Execute				:= bHomeAxis,
	Reset				:= bReset,	// #155
	StopActive			:= bStopAxis OR ((axisRef.NcToPlc.StateDWord AND 16#20000000) <> 0),	// #113
	Direction 			:= MC_Home_Direction.mcPositiveDirection,
	Velocity 			:= 1.0,
	Acceleration		:= 3.6,
	Deceleration		:= 3.6,
	Jerk				:= 3.6,
	RefPosition			:= -15.61+1.8,
	RefDistance			:= 5.18,
	TimeLimit 			:= T#1M,
	DistanceLimit 		:= 6,
	TravelLimit			:= 21,	// #165: 3 steps of 6 deg and the 2 deg jog, plus a margin
	Error 				=> bLatchHomeError,
	ErrorID 			=> nLatchHomeErrorID);
	


// #198
bSweepActive := bHomeAxis OR fbLatchHome.Busy;

// #69: FB_LatchHome clears its error as soon as Execute falls, and Execute falls on bError, so the error lasted
// one scan: the power-on was aborted, bError was FALSE again and no reset could fire. Hold it until the axis reset.
IF bReset THEN
	bLatchHomeErrorHeld := FALSE;
	nLatchHomeErrorIDHeld := 0;
END_IF
IF bLatchHomeError THEN
	bLatchHomeErrorHeld := TRUE;
	nLatchHomeErrorIDHeld := nLatchHomeErrorID;
END_IF

bError := bLatchHomeErrorHeld OR bAxisError;

// nErrorID is the current error: it used to keep stale values, so healthy axes were reset on every reset pass
IF bAxisError THEN
	nErrorID := nAxisErrorID;
ELSIF bLatchHomeErrorHeld THEN
	nErrorID := nLatchHomeErrorIDHeld;
ELSE
	nErrorID := 0;
END_IF
	
IF fbAxis.MoveDone OR bReset OR bError THEN
	bMoveAxis := FALSE;
END_IF

IF (fbAxis.HomeDone AND fbLatchHome.Done) OR bReset OR bError THEN
	bHomeAxis := FALSE;
END_IF
	
IF fbAxis.ResetDone THEN
	bReset := FALSE;
END_IF

// #159: bStopAxis was cleared only on StopDone. A stop of an axis that is disabled or standing still gives none, so
// it stayed TRUE and held every following sweep until a Reset Cold.
IF fbAxis.StopDone OR NOT bEnable OR bReset THEN
	bStopAxis := FALSE;
END_IF


bReady := fbAxis.Ready;

fbReadParameter(	
	Axis 			:= axisRef, 
	Enable 			:= fbAxis.InMotion, 
	ParameterNumber := MC_AxisParameter.AxisRemainingTimeToGo, 
	ReadMode 		:= E_ReadMode.READMODE_CYCLIC);
				
IF fbReadParameter.Valid THEN
	fSlewtime := fbReadParameter.Value;
END_IF


axisEvent(	
	Trigger 		:= bError, 
	Level 			:= ADSLOG_MSGTYPE_ERROR,
	FormatString	:= 'Declination Axis Error: %s',
	OnMessage 		:= NCError_TO_STRING(nErrorID),
	OffMEssage 		:= 'OK',
	OffLevel 		:= ADSLOG_MSGTYPE_HINT,
	Comm			:= fbComm);
	

CalibrationEvent(	
	Trigger 		:= bCalibrated, 
	Level 			:= ADSLOG_MSGTYPE_HINT,
	OnMessage 		:= 'Declination Axis is calibrated.',
	Comm			:= fbComm);

// Homing goes through FB_LatchHome and MC_SetPosition on bHomeAxis (the level), not through fbAxis.Home(), so this
// is empty (abstract in BROTLib's FB_BaseAxis, BROTLib #62).
METHOD _StartHoming : BOOL
_StartHoming := TRUE;
END_METHOD

END_FUNCTION_BLOCK

// ---- POUs/FB_TelescopeControl.TcPOU
FUNCTION_BLOCK FB_TelescopeControl EXTENDS BROTLib.FB_RaDecTelescopeControl
VAR_INPUT
(*
TCS interface section
see https://gitlab.aip.de/bmk10k/telescope_firmware/snippets/5
*)
	bSafetyAckRequest	: BOOL;		// set by a telescope reset, taken (and cleared) by MAIN which gives the safety acknowledge (#11)
	bStartupAxisReset	: BOOL;		// set by MAIN once when the safety start-up is done: one axis reset pass like after the reset acknowledge (#103)
	fPoleZone			: LREAL := 3.0;		// 90° - fPoleZone = No go zone near the Pole
	fPointingSafeAltitude	: LREAL := 5.0;	// ELEVATION below which the pointing model's fixed-point inversion is not numerically reliable (chaotic, see FB_PointingModelInversion / testing/check_pointing_inversion.py); gates goto/slew targets and tracking in addition to fHorizon
	
	fSlewVelocity		: LREAL := 8.0;		// Motor velocity for moving the telescope in degree/s
	
	// TRUE while the E-stop is triggered (MAIN: safetyHandling.estop): disables both axes, which only the next
	// power-on enables again, and publishes STATUS.GLOBAL = 1
	// MAIN: safetyHandling.ackPending (previous scan). An E-stop was seen and no clean safety acknowledge has run
	// since: the reset fires on it even without an error, and a power-on is refused (#59)
	bSafetyAckPending	: BOOL	:= FALSE;
    fStartupFocusTolerance : LREAL := 0.005; // match FB_FocusControl.fTolerance; align if that axis setting changes
	fbFocus				: I_Focus;
	fbCovers			: I_MirrorCovers;
	fbDome				: I_Dome;

	fbHourAngle			: REFERENCE TO FB_HourAngleControl;
	fbDeclination		: REFERENCE TO FB_DeclinationControl;

END_VAR
VAR
	fbCabinet			: FB_CabinetControl;

	fHourAnglePointingOffset	: LREAL; // pointing offset to sky
	fDeclinationPointingOffset	: LREAL; // pointing offset to sky
	fHourAngleInversionOffset	: LREAL;
	fDeclinationInversionOffset : LREAL;
	fHourAngleInversionOffsetCalc	: LREAL;	// raw output of fbPointingInversion this cycle, only copied into fHourAngleInversionOffset when bPointingInversionValid
	fDeclinationInversionOffsetCalc : LREAL;
	bPointingInversionValid		: BOOL;		// FALSE near the horizon where the inversion doesn't converge; fHourAngleInversionOffset/fDeclinationInversionOffset then keep their last valid value
	fHourAngleVelocity			: LREAL;	// rotational velocity of the HourAngle
	fDeclinationVelocity		: LREAL;	// rotational velocity of the Declination
	fbEq2Hor			: FB_EQ2HOR;
	fbHor2Eq			: FB_HOR2EQ;
	fbHaDec2RaDec		: FB_HADEC2RADEC;
	fbRaDec2HaDec		: FB_RADEC2HADEC;
	fbPointingForward	: FB_PointingModelForward;
	fbPointingInversion : FB_PointingModelInversion;
	
	bAxesCalibrated		: BOOL;		// #161: horizon/pole stops only act on a referenced counter
	bPowerOnHold		: BOOL;		// #166: a power-on is running and may be enabling a still axis inside a limit
	bHaMoving, bDecMoving	: BOOL;	// #166
	rtrigCalibLost		: F_TRIG;	// #161: calibration lost while enabled
	rtrigHorizonError	: R_TRIG;		// if the set Coordinate is below the Horizon threshold fHorizon
	rtrigPoleError		: R_TRIG;		// if the set Coordinate is in the pole zone fPoleZone
	
	rtrigResetAny		: R_TRIG;		// every reset edge (method, input, cabinet key), also without an error: the request part of the reset
	rtrigPoweredClear	: R_TRIG;		// #100: error or E-stop edge: the telescope is no longer powered
	bAxisResetAfterAck	: BOOL;		// reset the errored axes a second time once the acknowledge is done (#11)
	tonAxisResetAfterAck	: TON;
	// plan step 3.2: the axis feedback of this scan (1 hour angle, 2 declination), filled by _ReadAxes
	aAxis				: ARRAY[1..2] OF ST_AxisStatus;
	bHwErrorLast		: BOOL;		// BROTLib#25 step 4.4d: bHwError of the previous scan (edge for F_ErrorParkRequest)
	bErrorParkStarted	: BOOL;		// the park that a new axis/focus error starts (MONETcommon#86)
	bResetRequest		: BOOL;		// Reset() was called (one scan); kept apart from bResetActive, which the trigger below drives (#36)
	nSoftwareErrorID	: UDINT;	// 16#10 goto, 16#20 park, 16#30 home, 16#40 slew timeout
	bParkInError		: BOOL;		// a park was requested during an error (one scan): covers closed, dome parked, mount not moved
	sParkEnd			: STRING(160) := 'completed';	// the park log line when bParkActive falls: completed, or why it ended (#57)
	bParkLogged			: BOOL;		// bParkActive as the park event saw it last scan: PARK commencing is logged, an end line follows (#57)
	sParkWhy			: STRING(160);	// what the emergency park commanded, for the park log lines (#57)
	sHomeEnd			: STRING(40) := 'completed';	// the same for the home (#75)
	bHomeCancelled		: BOOL;		// a pending home that never started was dropped (one scan): logs the reason (#75)
	sHomeDropWhy		: STRING(160);	// why the pending home was dropped, for the WARN text (#108)
	fbStopTx			: BROTLib.FB_StopTransaction;	// #108/#120: one stop per axis and stop transaction
	rtHaMove			: R_TRIG;		// #92: MoveAxis of the axis went TRUE: the move command is out (MoveTo)
	rtDecMove			: R_TRIG;
	bHaMovePending		: BOOL;			// #92: a move was commanded and the NC does not report it yet: the axis is not at rest
	bDecMovePending		: BOOL;
	tonHaMovePending	: TON;			// #92: a command the NC never started (cancelled in time) is forgotten after 1 s
	tonDecMovePending	: TON;
	fbHomeDrop			: FB_HomeDropReason;	// #108/#120: why a pending home was dropped
	tonHomePending		: FB_TimeoutTimer;		// #75: bGoHome set but the home is not running (not ready, powered off): cancelled after 2 min
	
	bInitRefused		: BOOL;		// Init() was refused because of a stop or a park (one scan): logs 'power-on ignored: <reason>'
	sInitRefusedReason	: STRING(80);
	nInitRefusedCount	: UDINT;	// diagnostics (ADS)
	TCSinitRefusedEvent	: FB_Eventlog;
	bPowerBlocked		: BOOL;		// a power-on request was refused because of an error (one scan): logs the reason, every time
	bInHorizonLimit		: BOOL;		// #84: the mount is below the horizon limit (the safety block homes it out)
	bInPoleLimit		: BOOL;		// #84: the mount (or the tracking target) is in the pole zone
	bLimitHome			: BOOL;		// #84: the pending or running home was requested by a limit block; latched while bGoHome
	bParkAfterHome		: BOOL;		// #84: a park waits for that home
	bParkHomeDone		: BOOL;		// #84: the home finished for this park: the limit blocks do not home again, the park runs
	bParkHomeFirst		: BOOL;		// #84: a park was requested in a limit, the home runs first (one scan): logs it
	bSafeParked			: BOOL;		// an axes-off park is closing the covers and parking the dome, the mount was not moved: READY_STATE 0.3 until done (#110, #187)
	bParkedInPlace		: BOOL;		// the last park ended where the mount stood (axes off, covers closed, dome parked): bIsParked is TRUE, the mount may not be at the park position (#187)
	bStopIgnored		: BOOL;		// #196: a stop arrived during the in-place park (one scan): logs that it is ignored
	bParkInPlaceDone	: BOOL;		// an axes-off park just ended (one scan): logs it
	bParkInPlaceOpen	: BOOL;		// #197/#200: the park that logged PARK commencing goes on as an in-place park; its end line is the PARK end line
	sParkInPlaceEnd		: STRING(160);	// #200: how the in-place park ended: completed in place, or why it was aborted
	nParkInPlaceLevel	: DWORD := ADSLOG_MSGTYPE_HINT;
	tonParkPending		: FB_TimeoutTimer;		// #197: a park that is requested but never starts is forced into an in-place park after 2 min
	bParkForceInPlace	: BOOL;		// #197: the pending-park watchdog fired
	tonParkInPlace		: FB_TimeoutTimer;		// #187: an axes-off park gives up after 120 s if the covers or the dome do not finish
	bHomeByCommand		: BOOL;		// the running or pending home was requested by a Home() call or a bGoHome edge; the power-on's own home and the limit homes are not: a move replaces them (the old precedence), only a commanded home rejects moves (gohome_active)
	bCommandRejected	: BOOL;		// set by _NoteRejected, logged and cleared by the body (as MONETcommon, #83)
	eLastRejectedCommand	: E_TCSCommand;
	eLastRejectReason	: BROTLib.E_CommandRejectReason;
	nCommandRejectCount	: UDINT;	// diagnostics (ADS)
	sRejectMessage		: STRING(120);
	tonRejectRepeat		: TON;		// an identical rejection within 2 s is logged once (all are counted)
	eLoggedCommand		: E_TCSCommand;
	eLoggedReason		: BROTLib.E_CommandRejectReason;
	sStopNoDone			: STRING(10);	// #120: the axes named in the stop timeout text
	bStopTimeoutLog		: BOOL;		// #120: the stop transaction timed out or was released by the timeout (one scan); text in TCSstopTimeoutEvent.OnMessage
	// MONETcommon#17: 600 s timeouts of the goto/home/slew state machines. They were TONs in the methods' plain VAR, which is
	// re-created on every call, so they never fired. Fed every scan in the body, reset when the command flag drops.
	tonGotoTimeout			: FB_TimeoutTimer;
	tonHomeTimeout			: FB_TimeoutTimer;
	tonSlewTimeout			: FB_TimeoutTimer;
	tonParkTimeout			: FB_TimeoutTimer;		// park had no state-machine timeout: covers that never close hung it forever
	tonParkFocus			: FB_TimeoutTimer;		// park stage 80 waits for the focus move to end (#56), at most 60 s
	
	TCSsoftErrorEvent,
	TCSparkErrorEvent,
	TCSparkInPlaceEvent,
	TCSstopIgnoredEvent,
	TCShomeCancelEvent,
	TCSpowerBlockedEvent,
	TCSpowerParkEvent,
	TCSparkHomeEvent		: FB_Eventlog;	// #30, park during an error, a blocked power-on (every request)
	RejectEvent				: FB_Eventlog;	// a move command that the acceptance table rejects (was TCScommandRefusedEvent, #100)
	TCSstopTimeoutEvent		: FB_Eventlog;	// #120: a stop transaction passed 30 s without a Done of an axis, and its release

	nStatusWord, nLastStatus:	UDINT;
	bTestError : BOOL; // Test Error, deactivates under reset command
END_VAR
VAR_OUTPUT
	bSliding			: BOOL;		//TRUE, IF telescope is in fast-MOVE phase (includes pole-swap)	
	fbSweepStop			: FB_SweepStop;	// #113: switches the uncalibrated axes off after a stop in the calibration sweep
	bSettled			: BOOL;		// #98: at rest AND no stop transaction running (every stopped axis reported Done, no motion lock): gate of every home/restart that follows a stop
	bLocalMode			: BOOL;		// TRUE if switch is flipped to prevent Robotic Mode
	// Request latches (BROTLib#25, IAG50cm command model step 1a): the command inputs bPower/bPark/bStop/bReset are edge-triggered and
	// never written by the block; these latches are the block's own state, set by Init()/Park()/Stop()/the reset trigger, cleared by the body
END_VAR
VAR CONSTANT
	fSiderialVelocity: LREAL := 360.0 / 86164.099;
END_VAR

// The command model is in FB_BaseTelescopeControl (BROTLib 0.20.0, #25 step 5.4); this block fills in its hook methods.
SUPER^();

// Hook of the template body (BROTLib#25 step 5.4, S3: the body of this block is the template text, the differences are in these methods). Start of the scan after the startup scan.
METHOD PROTECTED _ScanBegin
// nothing
END_METHOD

// Hook of the template body (BROTLib#25 step 5.4, S3: the body of this block is the template text, the differences are in these methods). Reads the inputs of the axes and the cabinet.
METHOD PROTECTED _ReadInputs
_ReadAxes();
// State of the Cabinet
fbCabinet(bEstop := bEstopTriggered, bSafetyAckPending := bSafetyAckPending);	// #93: error LED during E-stop / pending acknowledge
bLocalMode := fbCabinet.LocalMode;
END_METHOD

// Hook of the template body (BROTLib#25 step 5.4, S3: the body of this block is the template text, the differences are in these methods). Error ID, axis resets, slew time and the error flag of this scan.
METHOD PROTECTED _ReadErrors
// get error ID
IF fbHourAngle.Error THEN
	nErrorID := fbHourAngle.nErrorID;
ELSIF fbDeclination.bError THEN
	nErrorID := fbDeclination.nErrorID;
ELSIF fbFocus <> 0 AND_THEN fbFocus.Error THEN
	nErrorID := fbFocus.ErrorID;
ELSIF bSoftwareError THEN
	nErrorID := nSoftwareErrorID;
END_IF

// reset (#11): every errored axis in one go, not only the first one. The drives stay in STO until the safety
// acknowledge (MAIN, bSafetyAckRequest: ErrAck 1 s, Restart 1 s), so the axes are reset again once it is done.
// The second pass resets every axis that is errored or not enabled (#55): after an E-stop HA and Dec can have lost
// their enable without latching an error, and then failed at the next power-on (18000) until they got a reset.
// #103: the safety start-up (MAIN) acknowledges like the reset does, but nothing reset the axes afterwards. After a
// Reset Cold the first enable then failed with 18000 until a reset=1 gave the second pass below. Experiment: run that
// pass once after the start-up. It also holds the power-on at stages 0 and 40 for its 2.5 s, like after a reset.
IF bStartupAxisReset THEN
	bStartupAxisReset := FALSE;
	bAxisResetAfterAck := TRUE;
END_IF
IF bResetActive THEN
	bSafetyAckRequest := TRUE;
	bAxisResetAfterAck := TRUE;
	_ResetErroredAxes(bAll := FALSE);
END_IF
tonAxisResetAfterAck(IN := bAxisResetAfterAck, PT := T#2500MS);
IF tonAxisResetAfterAck.Q THEN
	bAxisResetAfterAck := FALSE;
	_ResetErroredAxes(bAll := TRUE);
END_IF

// fSlewTime
fSlewTime := fbHourAngle.fSlewTime + fbDeclination.fSlewTime;

// ERROR (either one of the Axis or below safe Horizon (fHorizon))
bError := fbHourAngle.Error OR fbDeclination.Error OR(fbFocus <> 0 AND_THEN fbFocus.Error) OR fbCabinet.Error OR bTestError OR bSoftwareError;
END_METHOD

// Hook of the template body (BROTLib#25 step 5.4, S3: the body of this block is the template text, the differences are in these methods). The reaction to an error before the move gate.
METHOD PROTECTED _ErrorReaction
// #100: an error or an E-stop ends the powered state. Only a power-on or a park wrote bIsPowered, so it stayed TRUE and the
// next power=1 could be taken for a running telescope. bReady needs bIsPowered, so this only forces the full power-on.
rtrigPoweredClear(CLK := bError OR bEstopTriggered);
IF rtrigPoweredClear.Q THEN
	bIsPowered := FALSE;
END_IF
END_METHOD

// Hook of the template body (BROTLib#25 step 5.4, S3: the body of this block is the template text, the differences are in these methods). A move input edge was accepted.
METHOD PROTECTED _OnMoveEdgeAccepted
VAR_INPUT
	eCommand	: E_TCSCommand;
END_VAR
// nothing
END_METHOD

// Hook of the template body (BROTLib#25 step 5.4, S3: the body of this block is the template text, the differences are in these methods). The axes and the cabinet LED on an error.
METHOD PROTECTED _ApplyError
IF bError THEN
	fbHourAngle.Enable := FALSE;
	fbDeclination.Enable := FALSE;
	fbCabinet.Error := TRUE;
ELSE
	fbCabinet.Error := FALSE;
END_IF
END_METHOD

// Hook of the template body (BROTLib#25 step 5.4, S3: the body of this block is the template text, the differences are in these methods). The target of this scan and the reported position.
METHOD PROTECTED _ComputeTargets
// calculate fHourAngleApparent, fDeclinationApparent 

fbRaDec2HaDec(
	ra := fRightAscension,
	dec := fDeclination,
	lon := telescopeConfig.longitude,
	JD := fJd + fTimeOffset,
	ha_out => fHourAngleApparent,
	dec_out => fDeclinationApparent);
// (and also horizontal coord. -> used for checking if target is on sky or in ground)
fbEq2Hor(
	ra := fRightAscension,
	dec := fDeclination,
	lon := telescopeConfig.longitude,
	lat := telescopeConfig.latitude,
	altitude := telescopeConfig.altitude,
	JD := fJd + fTimeOffset,
	refract_to_observed := TRUE,
	alt => fElevationCalc,
	az => fAzimuthCalc);
	
